// TIA Portal project "TestFineModuloPLC2SnideroEmanuele" (V19)

(* hardware
DEVICE "S7-1200 station_1"  S7-1200 Station
   slot 0: "Telaio di montaggio_0"  S7-1200 Rack  Rack  V1.0
   slot 1: "PLC_1"  CPU 1212C DC/DC/Rly  6ES7 212-1HE40-0XB0  V4.6
   slot 2: "DI 8/DQ 8x24VDC_1"  6ES7 223-1BH32-0XB0  V2.0
DEVICE "HMI_1"  KTP900 Basic PN
   slot 0: "HMI_1"  KTP900 Basic PN  6AV2 123-2JB03-0AX0  17.0.0.0
   slot 1: "HMI_RT_1"  KTP900 Basic PN  6AV2 123-2JB03-0AX0  17.0.0.0
   slot 5: "HMI_1.IE_CP_1"  PROFINET Interface  17.0.0.0
      slot 1: "Interfaccia_1 PROFINET"  PROFINET Interface
         slot 1: "Porta_1"  Port
DEVICE "SINAMICS G_1"  Sinamics.Device
   slot 0: "	_0"  Rail  SinamicsG120CRackP
   slot 0: "Drive_1"  G120C PN  6SL3210-1KE11-8AF2  4.7.14
      slot 1: "PROFINET interface"  MDD-SinamicsG120-P
      slot 3: "PM G120C"  PM G120C  6SL3210-1KE11-8AF2  -
*)

// ===== PLC "PLC_1"  CPU 1212C DC/DC/Rly =====

VAR_GLOBAL   // PLC tag table "Tabella delle variabili standard"
   "AbilitazioneAvvioNastro1" AT %I0.0 : Bool;
   "AbilitazioneAvvioNastro2" AT %I0.1 : Bool;
   "AbilitazioneAvvioNastro3" AT %I0.2 : Bool;
   "ArrestoNastro1" AT %I0.3 : Bool;
   "ArrestoNastro2" AT %I0.4 : Bool;
   "ArrestoNastro3" AT %I0.5 : Bool;
   "Emergenza" AT %I0.6 : Bool;
   "P01" AT %I0.7 : Bool;
   "P02" AT %I1.0 : Bool;
   "P1" AT %I1.1 : Bool;
   "P2" AT %I1.2 : Bool;
   "MotoreRobot" AT %Q0.0 : Bool;
   "MotoreAperturaPinza" AT %Q0.4 : Bool;
   "LEDLavorazione" AT %Q0.1 : Bool;
   "LEDRiposo" AT %Q0.2 : Bool;
   "LEDErrorePrelievoNastro1" AT %Q0.3 : Bool;
   "P03" AT %I1.4 : Bool;
   "P3" AT %I1.5 : Bool;
   "MotoreNastro1" AT %Q0.5 : Bool;
   "MotoreNastro2" AT %Q0.6 : Bool;
   "MotoreNastro3" AT %Q0.7 : Bool;
   "MotoreChiusuraPinza" AT %Q1.0 : Bool;
   "LEDErrorePrelievoNastro2" AT %Q1.1 : Bool;
   "Axis_1_Drive_IN" AT %I256.0 : "PD_TEL1_IN";
   "Axis_1_Drive_OUT" AT %Q256.0 : "PD_TEL1_OUT";
END_VAR

VAR_GLOBAL   // PLC tag table "Segnalazioni"
   "IndiceSegnalazioni" AT %MW100 : Int;
   "ErrorePrelievoNastro1" AT %M101.0 : Bool;
   "ErrorePrelievoNastro2" AT %M101.1 : Bool;
END_VAR

DATA_BLOCK "Sistema"   // DB1
{ S7_Optimized_Access := 'TRUE' }
VERSION : 0.1
   VAR
      DurataTrasportoNastri : Time := T#2500ms;
      DurataSpostamentoRobot : Time := T#2000ms;
      DurataMovimentoPinza : Time := T#2000ms;
      DurataPrelievoScatola : Time := T#20000ms;
      VolumeScatola : SInt := 6;
   END_VAR
   VAR RETAIN
      RiempimentoScatola : SInt;
   END_VAR
   VAR
      PP01 : Bool;
      PP02 : Bool;
      PP03 : Bool;
      PP1 : Bool;
      PP2 : Bool;
      PP3 : Bool;
      NMotoreNastro1 : Bool;
      NMotoreNastro2 : Bool;
      NMotoreNastro3 : Bool;
      NQTPSostituzioneScatola : Bool;
   END_VAR
   VAR RETAIN
      P1 : Bool;
      P2 : Bool;
   END_VAR
   VAR
      P3 : Bool;
      P03 : Bool;
      PP03Sistema : Bool;
      SetpointVelocitàNormato : Real;
   END_VAR
   VAR RETAIN
      SetpointVelocitàScalato : Real;
   END_VAR
BEGIN
END_DATA_BLOCK

DATA_BLOCK "HMI"   // DB4
{ S7_Optimized_Access := 'TRUE' }
VERSION : 0.1
   VAR
      StartNastro1 : Bool;
      StartNastro2 : Bool;
      StartNastro3 : Bool;
   END_VAR
   VAR RETAIN
      StopNastro1 : Bool := true;
      StopNastro2 : Bool := true;
      StopNastro3 : Bool := true;
      Emergenza : Bool;
   END_VAR
   VAR
      DitoFotocellulaNastro1 : Bool;
      DitoFotocellulaNastro2 : Bool;
      CaricamentoPezzoNastro1 : Bool;
      PCaricamentoPezzoNastro1 : Bool;
      CaricamentoPezzoNastro2 : Bool;
      PCaricamentoPezzoNastro2 : Bool;
   END_VAR
   VAR RETAIN
      Posizione1PinzaAperta : Bool;
      Posizione2PinzaAperta : Bool;
      Posizione3PinzaAperta : Bool;
      Posizione1PinzaChiusa : Bool;
      Posizione2PinzaChiusa : Bool;
      Posizione3PinzaChiusa : Bool;
      IndiceRicetta : Int := 1;
      NomeSetDati : String := 'Veloce';
   END_VAR
   VAR
      VisibilitàPezzoNastro1Veloce : Bool;
      VisibilitàPezzoNastro1Lento : Bool;
      VisibilitàPezzoNastro2Veloce : Bool;
      VisibilitàPezzoNastro2Lento : Bool;
      VisibilitàPezzoNastro3Veloce : Bool;
      VisibilitàPezzoNastro3Lento : Bool;
      SetpointVelocitàMotoreNastri : Real;
      VelocitàAttualeMotoreNastri : Real;
   END_VAR
BEGIN
END_DATA_BLOCK

DATA_BLOCK "Robot_DB"   // DB6
{ S7_Optimized_Access := 'TRUE' }
VERSION : 0.1
// stored: InstanceOfName Robot
"Robot"
BEGIN
END_DATA_BLOCK

DATA_BLOCK "SetDatiSistema"   // DB9
{ S7_Optimized_Access := 'TRUE' }
VERSION : 0.1
   VAR
      DurataTrasportoNastri : Time := T#5000ms;
      DurataSpostamentoRobot : Time := T#4000ms;
      VolumeScatola : SInt := 3;
   END_VAR
BEGIN
END_DATA_BLOCK

DATA_BLOCK "SetDatiSistemaVeloce"   // DB10
{ S7_Optimized_Access := 'TRUE' }
VERSION : 0.1
   VAR
      DurataTrasportoNastri : Time := T#5000ms;
      DurataSpostamentoRobot : Time := T#4000ms;
      VolumeScatola : SInt := 3;
   END_VAR
BEGIN
END_DATA_BLOCK

DATA_BLOCK "SetDatiSistemaLento"   // DB11
{ S7_Optimized_Access := 'TRUE' }
VERSION : 0.1
   VAR
      DurataTrasportoNastri : Time := T#5000ms;
      DurataSpostamentoRobot : Time := T#4000ms;
      VolumeScatola : SInt := 3;
   END_VAR
BEGIN
END_DATA_BLOCK

// folder: System blocks/Program resources

DATA_BLOCK "TPNastro1"   // DB2
{ S7_Optimized_Access := 'TRUE' }
AUTHOR : Simatic
FAMILY : IEC
NAME : IEC_TMR
VERSION : 1.0
// stored: InstanceOfName IEC_TIMER
"IEC_TIMER"
BEGIN
END_DATA_BLOCK

DATA_BLOCK "TPNastro2"   // DB3
{ S7_Optimized_Access := 'TRUE' }
AUTHOR : Simatic
FAMILY : IEC
NAME : IEC_TMR
VERSION : 1.0
// stored: InstanceOfName IEC_TIMER
"IEC_TIMER"
BEGIN
END_DATA_BLOCK

DATA_BLOCK "TPNastro3"   // DB5
{ S7_Optimized_Access := 'TRUE' }
AUTHOR : Simatic
FAMILY : IEC
NAME : IEC_TMR
VERSION : 1.0
// stored: InstanceOfName IEC_TIMER
"IEC_TIMER"
BEGIN
END_DATA_BLOCK

DATA_BLOCK "TPSostituzioneScatola"   // DB7
{ S7_Optimized_Access := 'TRUE' }
AUTHOR : Simatic
FAMILY : IEC
NAME : IEC_TMR
VERSION : 1.0
// stored: InstanceOfName IEC_TIMER
"IEC_TIMER"
BEGIN
END_DATA_BLOCK

// folder: (top level)

DATA_BLOCK "Axis_1"   // DB12, Motion_DB
{ S7_Optimized_Access := 'TRUE' }
AUTHOR : SIMATIC
FAMILY : BasicMC
NAME : TO_PosAx
VERSION : 8.0
// stored: InstanceOfName TO_PositioningAxis
"TO_PositioningAxis"
BEGIN
   // Axis.Drive.OfflineDataAdaption = TRUE
   // Axis.Drive.TelegramAddressOutCU = %Q256.0
   // Axis.Drive.TelegramAddressInCU = %I256.0
   // Axis.Drive.DoNameCU = Drive_1.Standard_telegram_1
   // Axis.Encoder.SelectedHscIndexCU = -1
   // Axis.LengthUnitNormalized.Time = 1
   // Axis.LengthUnitNormalized.Distance = -2
   // Axis.Encoder.DbTypeCU = Classic
   // Axis.Drive.DbTypeCU = Classic
END_DATA_BLOCK

FUNCTION_BLOCK "Robot"   // FB1, LAD
{ S7_Optimized_Access := 'TRUE' }
VERSION : 0.1
   VAR_INPUT
      Obiettivo : SInt;   // 0 = HOME, 1 = OK1, 2 = OK2, 3 = OK3
   END_VAR
   VAR RETAIN
      PosizioneAttuale : SInt;   // 0 = HOME, 1 = OK1, 2 = OK2, 3 = OK3
      PinzaAperta : Bool := true;
      PezzoPrelevatoDaNastro1 : Bool;
      PezzoPrelevatoDaNastro2 : Bool;
   END_VAR
   VAR
      TPRotazioneRobot : TP_TIME;
      NMotoreRobot : Bool;
      ObiettivoInRaggiungimento : SInt;
      PQTPRotazioneRobot : Bool;
      TPPinza : TP_TIME;
      NTPRotazioneRobot : Bool;
      NMotoreChiusuraPinza : Bool;
      NMotoreAperturaPinza : Bool;
      BloccoRotazione : Bool;
   END_VAR
   VAR_TEMP   // added for the SCL form of the ladder/FBD networks
      _w1 : Bool;
      _w2 : Bool;
      _w3 : Bool;
      _w4 : Bool;
      _w5 : Bool;
      _w6 : Bool;
      _w7 : Bool;
      _w8 : Bool;
   END_VAR
BEGIN

REGION Network 1
   // ROTAZIONE BRACCIO e APERTURA/CHIUSURA PINZA
   // 
   // L'input di posizione obiettivo può cambiare durante lo spostamento del robot, ma ciò non influisce sulla meta in raggiungimento.
   // Va però salvata la posizione in raggiugimento per la durata dello spostamento.
   // 
   // Prima di muovere verso la prossima posizione bisogna attendere eventuali manovre di pinza (a meno che non ci si trovi in HOME)
   // 
   // La pinza è inizialmente aperta e resta aperta dopo il deposito sul nastro 3
   // 
   // Le fotocellule di fine corsa dei nastri 1 e 2 vengono resettate automaticamente a fine operazione di prelievo. L'errore è simulabile tramite PLCSIM o apposito pulsante HMI.
   // 
   // Può accadere che venga premuto il pulsante di emergenza durante il movimento: in tal caso si arrestano i motori e, al termine dello scorrimento del tempo previsto per i loro azionamenti, si resetta il blocco rotativo
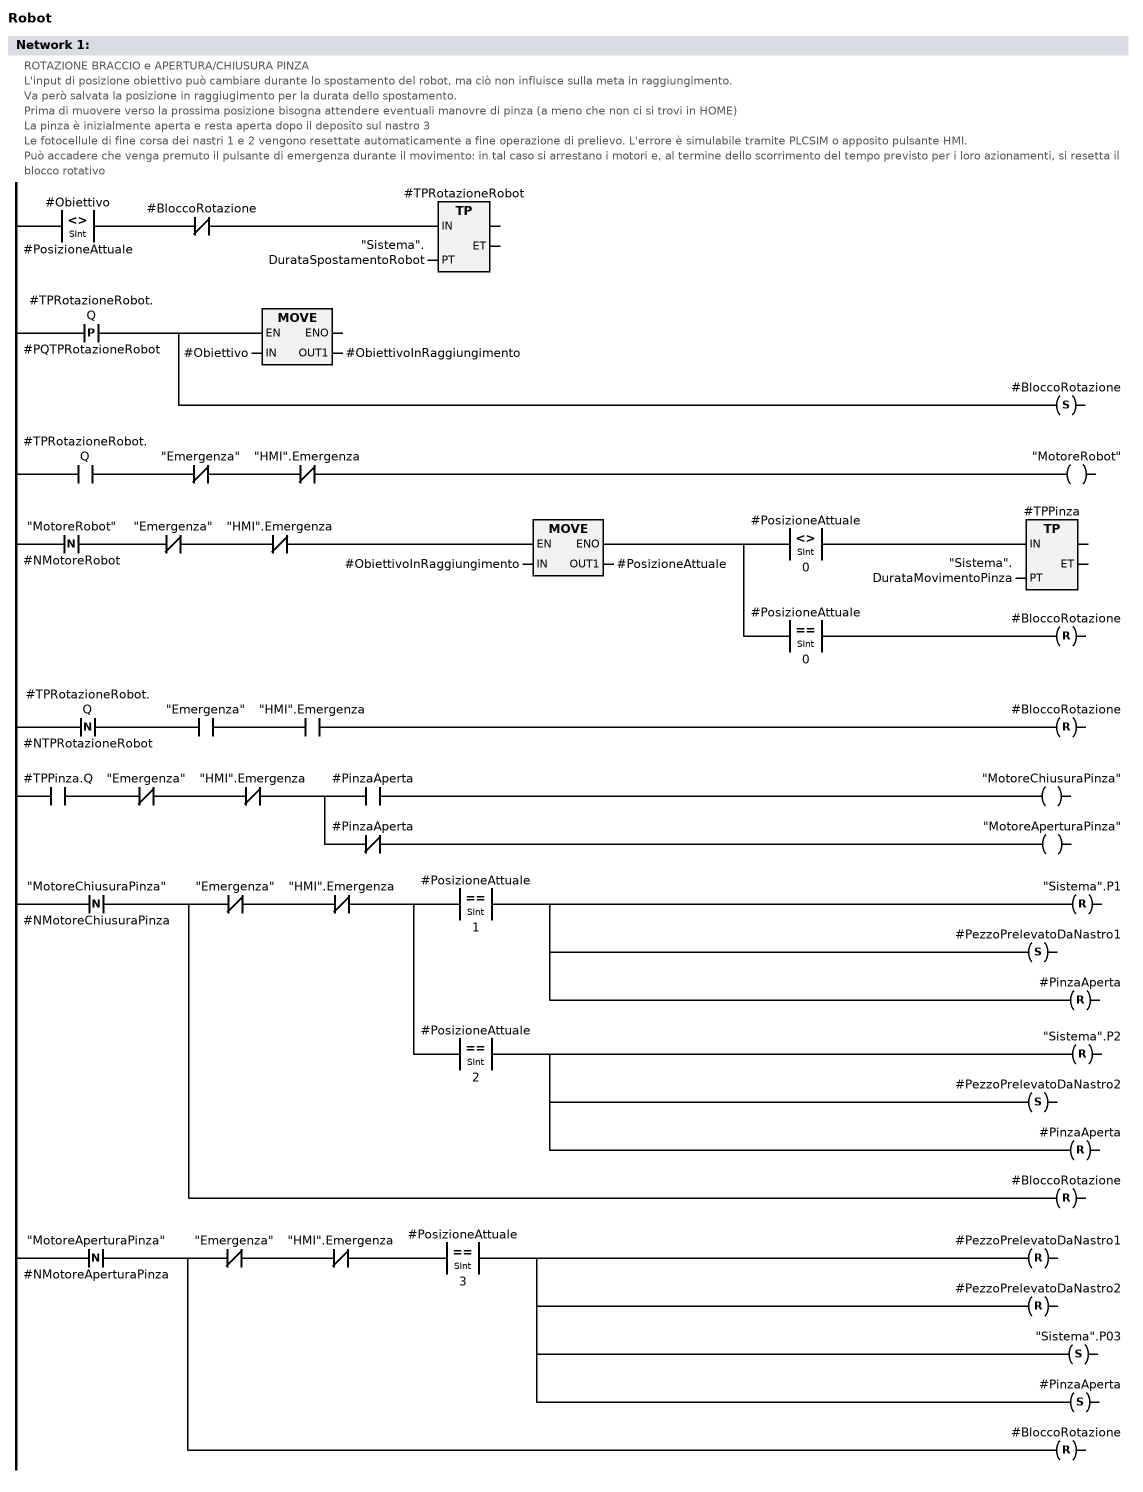
   #TPRotazioneRobot(IN := (#Obiettivo <> #PosizioneAttuale) AND NOT #BloccoRotazione,   // TP
                     PT := "Sistema".DurataSpostamentoRobot);
   #_w1 := #TPRotazioneRobot.Q AND NOT #PQTPRotazioneRobot;   // rising edge of #TPRotazioneRobot.Q
   #PQTPRotazioneRobot := #TPRotazioneRobot.Q;
   IF #_w1 THEN
       #ObiettivoInRaggiungimento := #Obiettivo;
       #BloccoRotazione := TRUE;
   END_IF;
   "MotoreRobot" := #TPRotazioneRobot.Q AND NOT "Emergenza" AND NOT "HMI".Emergenza;
   #_w2 := NOT "MotoreRobot" AND #NMotoreRobot;   // falling edge of "MotoreRobot"
   #NMotoreRobot := "MotoreRobot";
   #_w3 := #_w2 AND NOT "Emergenza" AND NOT "HMI".Emergenza;
   IF #_w3 THEN #PosizioneAttuale := #ObiettivoInRaggiungimento; END_IF;
   #TPPinza(IN := #_w3 AND (#PosizioneAttuale <> 0), PT := "Sistema".DurataMovimentoPinza);   // TP
   IF #_w3 AND (#PosizioneAttuale = 0) THEN #BloccoRotazione := FALSE; END_IF;
   #_w4 := NOT #TPRotazioneRobot.Q AND #NTPRotazioneRobot;   // falling edge of #TPRotazioneRobot.Q
   #NTPRotazioneRobot := #TPRotazioneRobot.Q;
   IF #_w4 AND "Emergenza" AND "HMI".Emergenza THEN #BloccoRotazione := FALSE; END_IF;
   #_w5 := #TPPinza.Q AND NOT "Emergenza" AND NOT "HMI".Emergenza;
   "MotoreChiusuraPinza" := #_w5 AND #PinzaAperta;
   "MotoreAperturaPinza" := #_w5 AND NOT #PinzaAperta;
   #_w6 := NOT "MotoreChiusuraPinza" AND #NMotoreChiusuraPinza;   // falling edge of "MotoreChiusuraPinza"
   #NMotoreChiusuraPinza := "MotoreChiusuraPinza";
   #_w7 := #_w6 AND NOT "Emergenza" AND NOT "HMI".Emergenza;
   IF #_w7 AND (#PosizioneAttuale = 1) THEN
       "Sistema".P1 := FALSE;
       #PezzoPrelevatoDaNastro1 := TRUE;
       #PinzaAperta := FALSE;
   END_IF;
   IF #_w7 AND (#PosizioneAttuale = 2) THEN
       "Sistema".P2 := FALSE;
       #PezzoPrelevatoDaNastro2 := TRUE;
       #PinzaAperta := FALSE;
   END_IF;
   IF #_w6 THEN #BloccoRotazione := FALSE; END_IF;
   #_w8 := NOT "MotoreAperturaPinza" AND #NMotoreAperturaPinza;   // falling edge of "MotoreAperturaPinza"
   #NMotoreAperturaPinza := "MotoreAperturaPinza";
   IF #_w8 AND NOT "Emergenza" AND NOT "HMI".Emergenza AND (#PosizioneAttuale = 3) THEN
       #PezzoPrelevatoDaNastro1 := FALSE;
       #PezzoPrelevatoDaNastro2 := FALSE;
       "Sistema".P03 := TRUE;
       #PinzaAperta := TRUE;
   END_IF;
   IF #_w8 THEN #BloccoRotazione := FALSE; END_IF;
END_REGION
END_FUNCTION_BLOCK

FUNCTION "AggiornamentoParametriRicetta" : Void   // FC2, LAD
{ S7_Optimized_Access := 'TRUE' }
VERSION : 0.1
   VAR_TEMP   // added for the SCL form of the ladder/FBD networks
      _w1 : Bool;
   END_VAR
BEGIN

REGION Network 1
   // Indice ricetta Sistema = 1
   // Indice salvato in Reciper Tag e in Data Record (HMI > Connections > Area Pointers)
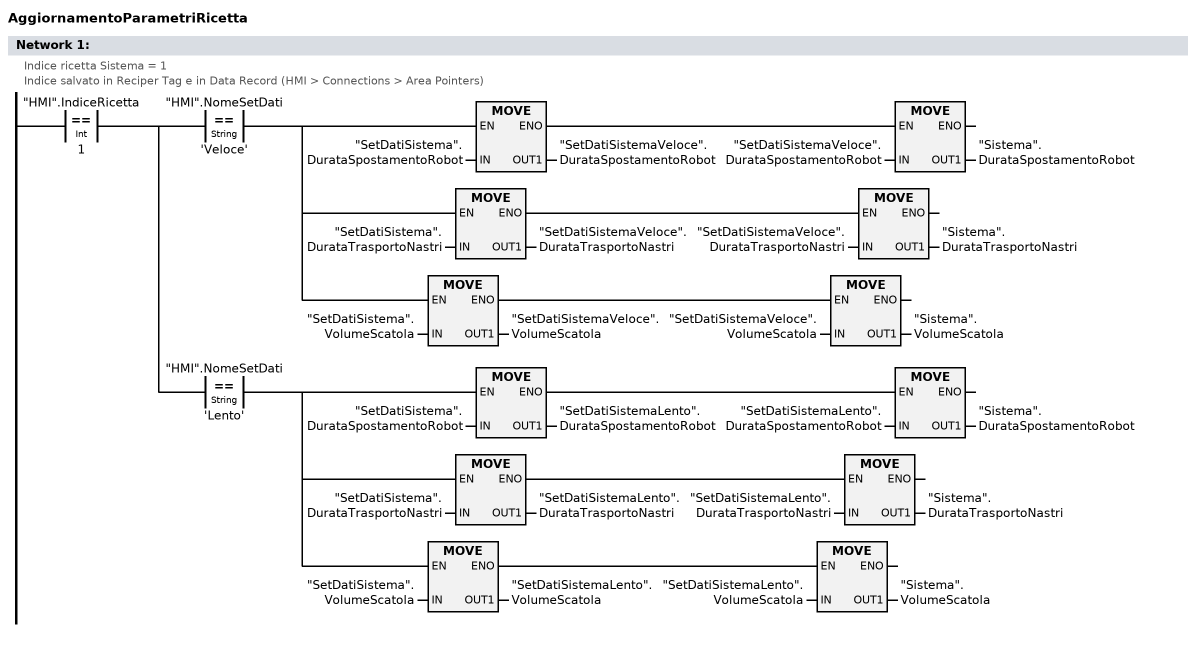
   RUNG wire#powerrail
      { S7_Templates := "SrcType := Int" } EQ_Contact(in1 := "HMI".IndiceRicetta, in2 := 1)
      wire#w1
      { S7_Templates := "SrcType := String" } EQ_Contact(in1 := "HMI".NomeSetDati, in2 := 'Veloce')
      wire#w2
      Move(in := "SetDatiSistema".DurataSpostamentoRobot, out1 => "SetDatiSistemaVeloce".DurataSpostamentoRobot)
      Move(in := "SetDatiSistemaVeloce".DurataSpostamentoRobot, out1 => "Sistema".DurataSpostamentoRobot)
   END_RUNG
   RUNG wire#w2
      Move(in := "SetDatiSistema".DurataTrasportoNastri, out1 => "SetDatiSistemaVeloce".DurataTrasportoNastri)
      Move(in := "SetDatiSistemaVeloce".DurataTrasportoNastri, out1 => "Sistema".DurataTrasportoNastri)
   END_RUNG
   RUNG wire#w2
      Move(in := "SetDatiSistema".VolumeScatola, out1 => "SetDatiSistemaVeloce".VolumeScatola)
      Move(in := "SetDatiSistemaVeloce".VolumeScatola, out1 => "Sistema".VolumeScatola)
   END_RUNG
   RUNG wire#w1
      { S7_Templates := "SrcType := String" } EQ_Contact(in1 := "HMI".NomeSetDati, in2 := 'Lento')
      wire#w3
      Move(in := "SetDatiSistema".DurataSpostamentoRobot, out1 => "SetDatiSistemaLento".DurataSpostamentoRobot)
      Move(in := "SetDatiSistemaLento".DurataSpostamentoRobot, out1 => "Sistema".DurataSpostamentoRobot)
   END_RUNG
   RUNG wire#w3
      Move(in := "SetDatiSistema".DurataTrasportoNastri, out1 => "SetDatiSistemaLento".DurataTrasportoNastri)
      Move(in := "SetDatiSistemaLento".DurataTrasportoNastri, out1 => "Sistema".DurataTrasportoNastri)
   END_RUNG
   RUNG wire#w3
      Move(in := "SetDatiSistema".VolumeScatola, out1 => "SetDatiSistemaLento".VolumeScatola)
      Move(in := "SetDatiSistemaLento".VolumeScatola, out1 => "Sistema".VolumeScatola)
   END_RUNG
   // the same network as SCL:
   #_w1 := "HMI".IndiceRicetta = 1;
   IF #_w1 AND ("HMI".NomeSetDati = 'Veloce') THEN
       "SetDatiSistemaVeloce".DurataSpostamentoRobot := "SetDatiSistema".DurataSpostamentoRobot;
       "Sistema".DurataSpostamentoRobot := "SetDatiSistemaVeloce".DurataSpostamentoRobot;
       "SetDatiSistemaVeloce".DurataTrasportoNastri := "SetDatiSistema".DurataTrasportoNastri;
       "Sistema".DurataTrasportoNastri := "SetDatiSistemaVeloce".DurataTrasportoNastri;
       "SetDatiSistemaVeloce".VolumeScatola := "SetDatiSistema".VolumeScatola;
       "Sistema".VolumeScatola := "SetDatiSistemaVeloce".VolumeScatola;
   END_IF;
   IF #_w1 AND ("HMI".NomeSetDati = 'Lento') THEN
       "SetDatiSistemaLento".DurataSpostamentoRobot := "SetDatiSistema".DurataSpostamentoRobot;
       "Sistema".DurataSpostamentoRobot := "SetDatiSistemaLento".DurataSpostamentoRobot;
       "SetDatiSistemaLento".DurataTrasportoNastri := "SetDatiSistema".DurataTrasportoNastri;
       "Sistema".DurataTrasportoNastri := "SetDatiSistemaLento".DurataTrasportoNastri;
       "SetDatiSistemaLento".VolumeScatola := "SetDatiSistema".VolumeScatola;
       "Sistema".VolumeScatola := "SetDatiSistemaLento".VolumeScatola;
   END_IF;
END_REGION
END_FUNCTION

ORGANIZATION_BLOCK "Main"   // OB1, LAD, ProgramCycle
TITLE = "Main Program Sweep (Cycle)"
{ S7_Optimized_Access := 'TRUE' }
VERSION : 0.1
   VAR_INPUT
      Initial_Call : Bool;   // Initial call of this OB
      Remanence : Bool;   // =True, if remanent data are available
   END_VAR
   VAR_TEMP   // added for the SCL form of the ladder/FBD networks
      _w1 : Bool;
      _w2 : Bool;
      _w3 : Bool;
      _w4 : Bool;
   END_VAR
BEGIN

REGION Network 1
   // Trasporto pezzi nastro 1
   // 
   // Non è possibile posizionare pezzi sui nastri finché ne sono in trasporto altri (o, meglio, è possibile ma il motore si fermerà si muoverà solamente per permettere) o la fotocellula di fine corsa non viene liberata (il motore non si aziona)
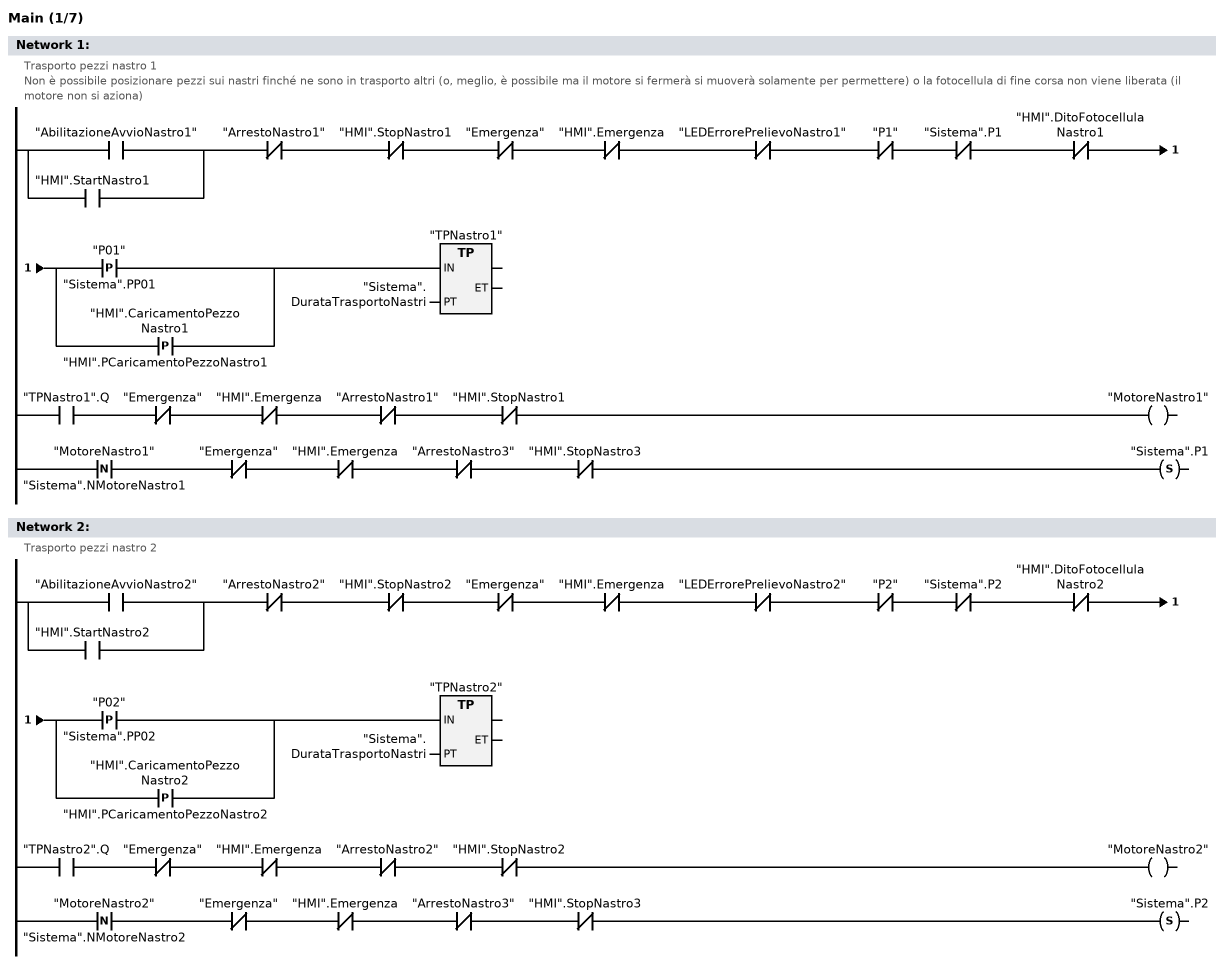
   #_w1 := ("AbilitazioneAvvioNastro1" OR "HMI".StartNastro1) AND NOT "ArrestoNastro1" AND NOT "HMI".StopNastro1 AND NOT "Emergenza" AND NOT "HMI".Emergenza AND NOT "LEDErrorePrelievoNastro1" AND NOT "P1" AND NOT "Sistema".P1 AND NOT "HMI".DitoFotocellulaNastro1 AND "P01" AND NOT "Sistema".PP01;   // rising edge of "P01"
   "Sistema".PP01 := "P01";
   #_w2 := ("AbilitazioneAvvioNastro1" OR "HMI".StartNastro1) AND NOT "ArrestoNastro1" AND NOT "HMI".StopNastro1 AND NOT "Emergenza" AND NOT "HMI".Emergenza AND NOT "LEDErrorePrelievoNastro1" AND NOT "P1" AND NOT "Sistema".P1 AND NOT "HMI".DitoFotocellulaNastro1 AND "HMI".CaricamentoPezzoNastro1 AND NOT "HMI".PCaricamentoPezzoNastro1;   // rising edge of "HMI".CaricamentoPezzoNastro1
   "HMI".PCaricamentoPezzoNastro1 := "HMI".CaricamentoPezzoNastro1;
   "TPNastro1".TP(IN := #_w1 OR #_w2, PT := "Sistema".DurataTrasportoNastri);
   "MotoreNastro1" := "TPNastro1".Q AND NOT "Emergenza" AND NOT "HMI".Emergenza AND NOT "ArrestoNastro1" AND NOT "HMI".StopNastro1;
   #_w3 := NOT "MotoreNastro1" AND "Sistema".NMotoreNastro1;   // falling edge of "MotoreNastro1"
   "Sistema".NMotoreNastro1 := "MotoreNastro1";
   IF #_w3 AND NOT "Emergenza" AND NOT "HMI".Emergenza AND NOT "ArrestoNastro3" AND NOT "HMI".StopNastro3 THEN
       "Sistema".P1 := TRUE;
   END_IF;
END_REGION

REGION Network 2
   // Trasporto pezzi nastro 2
   #_w1 := ("AbilitazioneAvvioNastro2" OR "HMI".StartNastro2) AND NOT "ArrestoNastro2" AND NOT "HMI".StopNastro2 AND NOT "Emergenza" AND NOT "HMI".Emergenza AND NOT "LEDErrorePrelievoNastro2" AND NOT "P2" AND NOT "Sistema".P2 AND NOT "HMI".DitoFotocellulaNastro2 AND "P02" AND NOT "Sistema".PP02;   // rising edge of "P02"
   "Sistema".PP02 := "P02";
   #_w2 := ("AbilitazioneAvvioNastro2" OR "HMI".StartNastro2) AND NOT "ArrestoNastro2" AND NOT "HMI".StopNastro2 AND NOT "Emergenza" AND NOT "HMI".Emergenza AND NOT "LEDErrorePrelievoNastro2" AND NOT "P2" AND NOT "Sistema".P2 AND NOT "HMI".DitoFotocellulaNastro2 AND "HMI".CaricamentoPezzoNastro2 AND NOT "HMI".PCaricamentoPezzoNastro2;   // rising edge of "HMI".CaricamentoPezzoNastro2
   "HMI".PCaricamentoPezzoNastro2 := "HMI".CaricamentoPezzoNastro2;
   "TPNastro2".TP(IN := #_w1 OR #_w2, PT := "Sistema".DurataTrasportoNastri);
   "MotoreNastro2" := "TPNastro2".Q AND NOT "Emergenza" AND NOT "HMI".Emergenza AND NOT "ArrestoNastro2" AND NOT "HMI".StopNastro2;
   #_w3 := NOT "MotoreNastro2" AND "Sistema".NMotoreNastro2;   // falling edge of "MotoreNastro2"
   "Sistema".NMotoreNastro2 := "MotoreNastro2";
   IF #_w3 AND NOT "Emergenza" AND NOT "HMI".Emergenza AND NOT "ArrestoNastro3" AND NOT "HMI".StopNastro3 THEN
       "Sistema".P2 := TRUE;
   END_IF;
END_REGION

REGION Network 3
   // Trasporto pezzi nastro 3 e riempimento scatola
   // 
   // Il nastro 3 non si muove se la scatola piena non è stata rimpiazzata
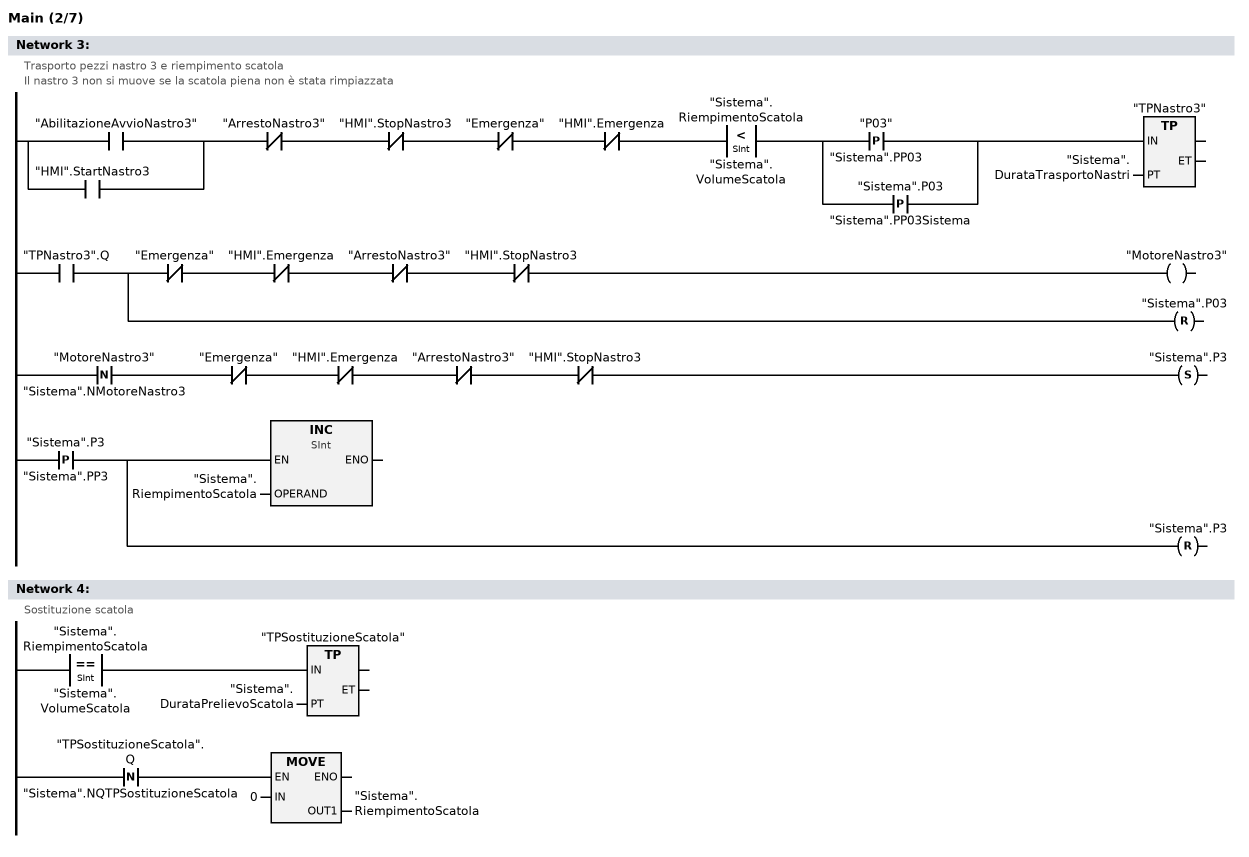
   #_w1 := ("AbilitazioneAvvioNastro3" OR "HMI".StartNastro3) AND NOT "ArrestoNastro3" AND NOT "HMI".StopNastro3 AND NOT "Emergenza" AND NOT "HMI".Emergenza AND ("Sistema".RiempimentoScatola < "Sistema".VolumeScatola) AND "P03" AND NOT "Sistema".PP03;   // rising edge of "P03"
   "Sistema".PP03 := "P03";
   #_w2 := ("AbilitazioneAvvioNastro3" OR "HMI".StartNastro3) AND NOT "ArrestoNastro3" AND NOT "HMI".StopNastro3 AND NOT "Emergenza" AND NOT "HMI".Emergenza AND ("Sistema".RiempimentoScatola < "Sistema".VolumeScatola) AND "Sistema".P03 AND NOT "Sistema".PP03Sistema;   // rising edge of "Sistema".P03
   "Sistema".PP03Sistema := "Sistema".P03;
   "TPNastro3".TP(IN := #_w1 OR #_w2, PT := "Sistema".DurataTrasportoNastri);
   "MotoreNastro3" := "TPNastro3".Q AND NOT "Emergenza" AND NOT "HMI".Emergenza AND NOT "ArrestoNastro3" AND NOT "HMI".StopNastro3;
   IF "TPNastro3".Q THEN "Sistema".P03 := FALSE; END_IF;
   #_w3 := NOT "MotoreNastro3" AND "Sistema".NMotoreNastro3;   // falling edge of "MotoreNastro3"
   "Sistema".NMotoreNastro3 := "MotoreNastro3";
   IF #_w3 AND NOT "Emergenza" AND NOT "HMI".Emergenza AND NOT "ArrestoNastro3" AND NOT "HMI".StopNastro3 THEN
       "Sistema".P3 := TRUE;
   END_IF;
   #_w4 := "Sistema".P3 AND NOT "Sistema".PP3;   // rising edge of "Sistema".P3
   "Sistema".PP3 := "Sistema".P3;
   IF #_w4 THEN
       "Sistema".RiempimentoScatola := "Sistema".RiempimentoScatola + 1;
       "Sistema".P3 := FALSE;
   END_IF;
END_REGION

REGION Network 4
   // Sostituzione scatola
   "TPSostituzioneScatola".TP(IN := "Sistema".RiempimentoScatola = "Sistema".VolumeScatola,
                           PT := "Sistema".DurataPrelievoScatola);
   #_w1 := NOT "TPSostituzioneScatola".Q AND "Sistema".NQTPSostituzioneScatola;   // falling edge of "TPSostituzioneScatola".Q
   "Sistema".NQTPSostituzioneScatola := "TPSostituzioneScatola".Q;
   IF #_w1 THEN "Sistema".RiempimentoScatola := 0; END_IF;
END_REGION

REGION Network 5
   // MOVIMENTAZIONE ROBOT
   // 
   // Spostamenti
   // - home => nastro 1/2
   // - nastro 1/2 => nastro 3
   // - nastro 3 => nastro1/2/home (se assenti pezzi da prelevare)
   // 
   // L'oggetto non viene prelevato per essere rilasciato sul nastro 3 finché il motore del nastro è in stato di arresto o la scatola è piena
   // Può però essere prelevato se il nastro 3 è in movimento perché vi è tempo sufficiente a completare l'inscatolamento del precedente prima che venga rilasciato.
   // 
   // Il nastro 1 ha precedenza sul 2
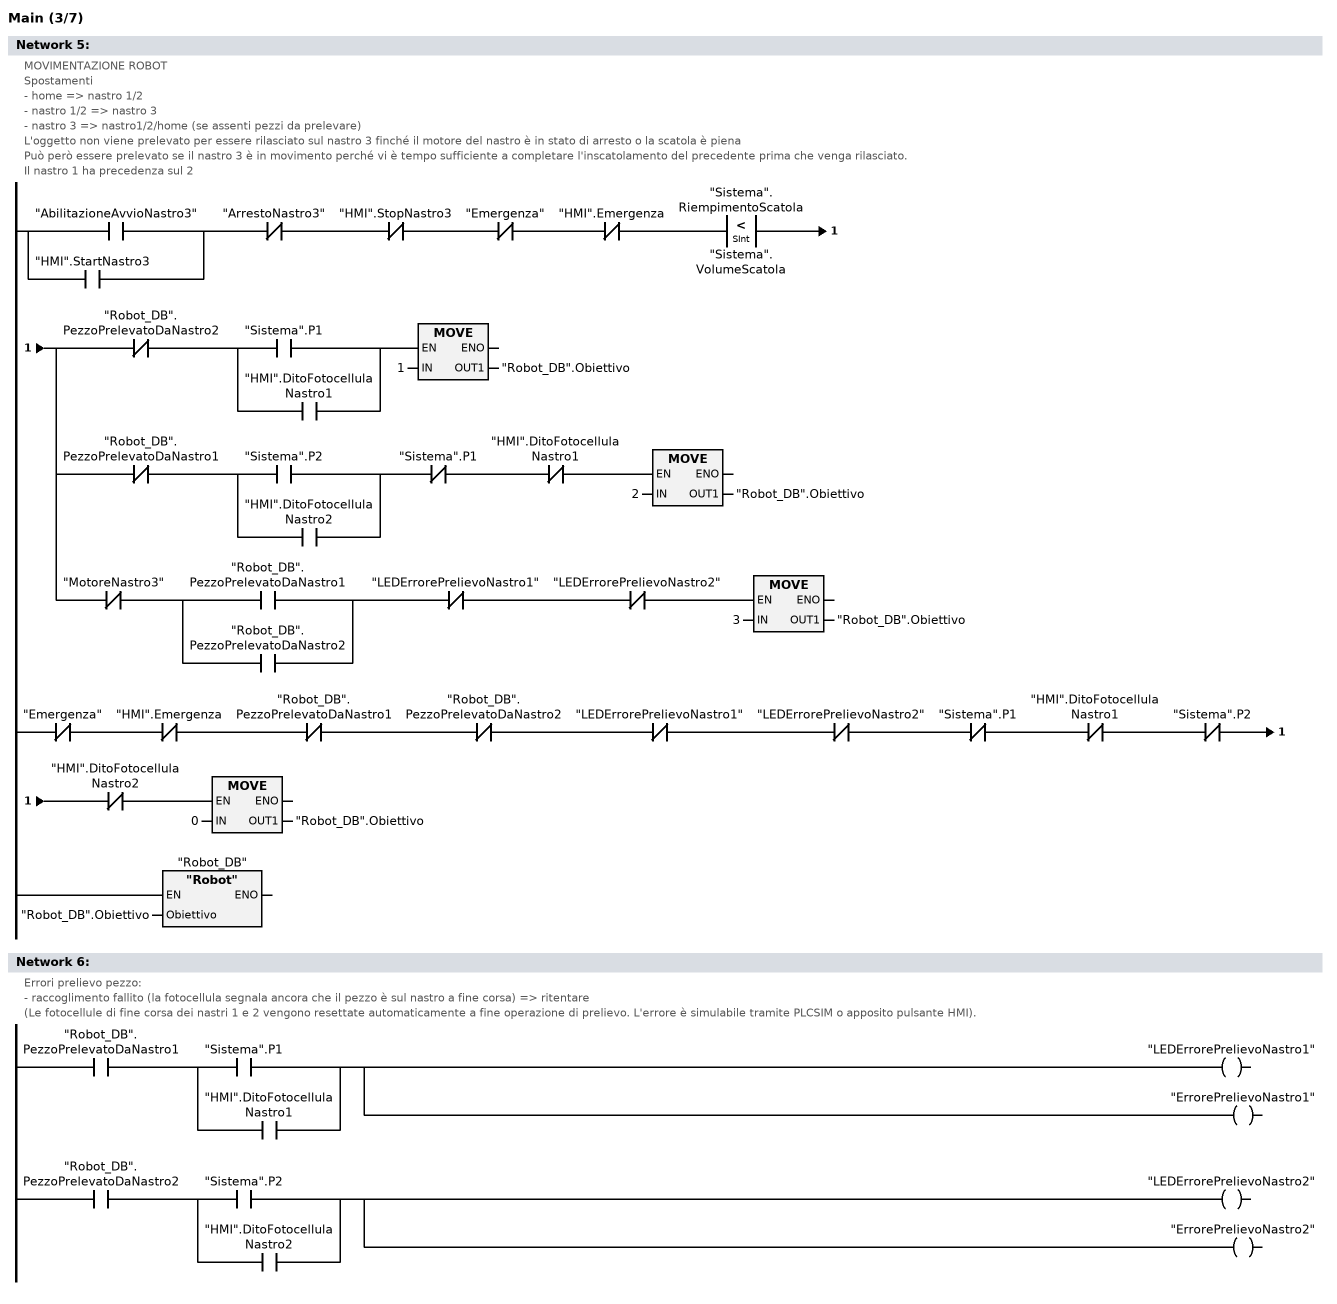
   RUNG wire#powerrail
      Contact( "AbilitazioneAvvioNastro3" )
      wire#w1
      I_Contact( "ArrestoNastro3" )
      I_Contact( "HMI".StopNastro3 )
      I_Contact( "Emergenza" )
      I_Contact( "HMI".Emergenza )
      { S7_Templates := "SrcType := SInt" } LT_Contact(in1 := "Sistema".RiempimentoScatola, in2 := "Sistema".VolumeScatola)
      wire#w2
      I_Contact( "Robot_DB".PezzoPrelevatoDaNastro2 )
      wire#w3
      Contact( "Sistema".P1 )
      wire#w4
      Move(in := 1, out1 => "Robot_DB".Obiettivo)
   END_RUNG
   RUNG wire#powerrail
      Contact( "HMI".StartNastro3 )
   END_RUNG wire#w1
   RUNG wire#w3
      Contact( "HMI".DitoFotocellulaNastro1 )
   END_RUNG wire#w4
   RUNG wire#w2
      I_Contact( "Robot_DB".PezzoPrelevatoDaNastro1 )
      wire#w5
      Contact( "Sistema".P2 )
      wire#w6
      I_Contact( "Sistema".P1 )
      I_Contact( "HMI".DitoFotocellulaNastro1 )
      Move(in := 2, out1 => "Robot_DB".Obiettivo)
   END_RUNG
   RUNG wire#w5
      Contact( "HMI".DitoFotocellulaNastro2 )
   END_RUNG wire#w6
   RUNG wire#w2
      I_Contact( "MotoreNastro3" )
      wire#w7
      Contact( "Robot_DB".PezzoPrelevatoDaNastro1 )
      wire#w8
      I_Contact( "LEDErrorePrelievoNastro1" )
      I_Contact( "LEDErrorePrelievoNastro2" )
      Move(in := 3, out1 => "Robot_DB".Obiettivo)
   END_RUNG
   RUNG wire#w7
      Contact( "Robot_DB".PezzoPrelevatoDaNastro2 )
   END_RUNG wire#w8
   RUNG wire#powerrail
      I_Contact( "Emergenza" )
      I_Contact( "HMI".Emergenza )
      I_Contact( "Robot_DB".PezzoPrelevatoDaNastro1 )
      I_Contact( "Robot_DB".PezzoPrelevatoDaNastro2 )
      I_Contact( "LEDErrorePrelievoNastro1" )
      I_Contact( "LEDErrorePrelievoNastro2" )
      I_Contact( "Sistema".P1 )
      I_Contact( "HMI".DitoFotocellulaNastro1 )
      I_Contact( "Sistema".P2 )
      I_Contact( "HMI".DitoFotocellulaNastro2 )
      Move(in := 0, out1 => "Robot_DB".Obiettivo)
   END_RUNG
   RUNG wire#powerrail
      "Robot_DB"(Obiettivo := "Robot_DB".Obiettivo)
   END_RUNG
   // the same network as SCL:
   #_w1 := ("AbilitazioneAvvioNastro3" OR "HMI".StartNastro3) AND NOT "ArrestoNastro3" AND NOT "HMI".StopNastro3 AND NOT "Emergenza" AND NOT "HMI".Emergenza AND ("Sistema".RiempimentoScatola < "Sistema".VolumeScatola);
   IF #_w1 AND NOT "Robot_DB".PezzoPrelevatoDaNastro2 AND ("Sistema".P1 OR "HMI".DitoFotocellulaNastro1) THEN
       "Robot_DB".Obiettivo := 1;
   END_IF;
   IF #_w1 AND NOT "Robot_DB".PezzoPrelevatoDaNastro1 AND ("Sistema".P2 OR "HMI".DitoFotocellulaNastro2) AND NOT "Sistema".P1 AND NOT "HMI".DitoFotocellulaNastro1 THEN
       "Robot_DB".Obiettivo := 2;
   END_IF;
   IF #_w1 AND NOT "MotoreNastro3" AND ("Robot_DB".PezzoPrelevatoDaNastro1 OR "Robot_DB".PezzoPrelevatoDaNastro2) AND NOT "LEDErrorePrelievoNastro1" AND NOT "LEDErrorePrelievoNastro2" THEN
       "Robot_DB".Obiettivo := 3;
   END_IF;
   IF NOT "Emergenza" AND NOT "HMI".Emergenza AND NOT "Robot_DB".PezzoPrelevatoDaNastro1 AND NOT "Robot_DB".PezzoPrelevatoDaNastro2 AND NOT "LEDErrorePrelievoNastro1" AND NOT "LEDErrorePrelievoNastro2" AND NOT "Sistema".P1 AND NOT "HMI".DitoFotocellulaNastro1 AND NOT "Sistema".P2 AND NOT "HMI".DitoFotocellulaNastro2 THEN
       "Robot_DB".Obiettivo := 0;
   END_IF;
   "Robot_DB"(Obiettivo := "Robot_DB".Obiettivo);   // "Robot"
END_REGION

REGION Network 6
   // Errori prelievo pezzo: 
   // - raccoglimento fallito (la fotocellula segnala ancora che il pezzo è sul nastro a fine corsa) => ritentare
   // 
   // (Le fotocellule di fine corsa dei nastri 1 e 2 vengono resettate automaticamente a fine operazione di prelievo. L'errore è simulabile tramite PLCSIM o apposito pulsante HMI).
   RUNG wire#powerrail
      Contact( "Robot_DB".PezzoPrelevatoDaNastro1 )
      wire#w1
      Contact( "Sistema".P1 )
      wire#w2
      Coil( "LEDErrorePrelievoNastro1" )
   END_RUNG
   RUNG wire#w1
      Contact( "HMI".DitoFotocellulaNastro1 )
   END_RUNG wire#w2
   RUNG wire#w2
      Coil( "ErrorePrelievoNastro1" )
   END_RUNG
   RUNG wire#powerrail
      Contact( "Robot_DB".PezzoPrelevatoDaNastro2 )
      wire#w3
      Contact( "Sistema".P2 )
      wire#w4
      Coil( "LEDErrorePrelievoNastro2" )
   END_RUNG
   RUNG wire#w3
      Contact( "HMI".DitoFotocellulaNastro2 )
   END_RUNG wire#w4
   RUNG wire#w4
      Coil( "ErrorePrelievoNastro2" )
   END_RUNG
   // the same network as SCL:
   "LEDErrorePrelievoNastro1" := "Robot_DB".PezzoPrelevatoDaNastro1 AND ("Sistema".P1 OR "HMI".DitoFotocellulaNastro1);
   "ErrorePrelievoNastro1" := "LEDErrorePrelievoNastro1";
   "LEDErrorePrelievoNastro2" := "Robot_DB".PezzoPrelevatoDaNastro2 AND ("Sistema".P2 OR "HMI".DitoFotocellulaNastro2);
   "ErrorePrelievoNastro2" := "LEDErrorePrelievoNastro2";
END_REGION

REGION Network 7
   // Alimentazione LED marcia sistema quando:
   // - il robot è in rotazione o in azionamento pinza
   // - un nastro è in scorrimento
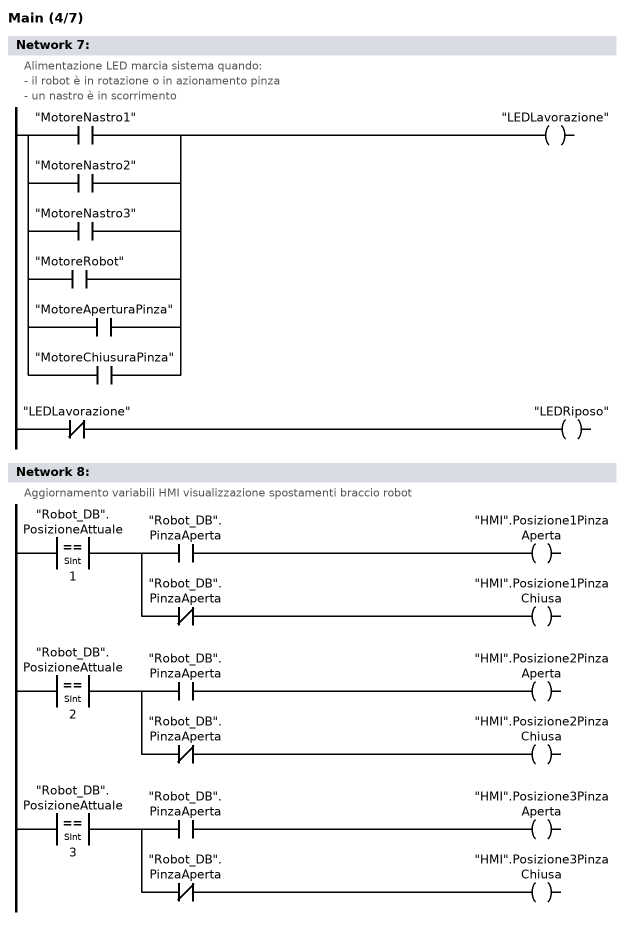
   RUNG wire#powerrail
      Contact( "MotoreNastro1" )
      wire#w1
      Coil( "LEDLavorazione" )
   END_RUNG
   RUNG wire#powerrail
      Contact( "MotoreNastro2" )
   END_RUNG wire#w1
   RUNG wire#powerrail
      Contact( "MotoreNastro3" )
   END_RUNG wire#w1
   RUNG wire#powerrail
      Contact( "MotoreRobot" )
   END_RUNG wire#w1
   RUNG wire#powerrail
      Contact( "MotoreAperturaPinza" )
   END_RUNG wire#w1
   RUNG wire#powerrail
      Contact( "MotoreChiusuraPinza" )
   END_RUNG wire#w1
   RUNG wire#powerrail
      I_Contact( "LEDLavorazione" )
      Coil( "LEDRiposo" )
   END_RUNG
   // the same network as SCL:
   "LEDLavorazione" := "MotoreNastro1" OR "MotoreNastro2" OR "MotoreNastro3" OR "MotoreRobot" OR "MotoreAperturaPinza" OR "MotoreChiusuraPinza";
   "LEDRiposo" := NOT "LEDLavorazione";
END_REGION

REGION Network 8
   // Aggiornamento variabili HMI visualizzazione spostamenti braccio robot
   RUNG wire#powerrail
      { S7_Templates := "SrcType := SInt" } EQ_Contact(in1 := "Robot_DB".PosizioneAttuale, in2 := 1)
      wire#w1
      Contact( "Robot_DB".PinzaAperta )
      Coil( "HMI".Posizione1PinzaAperta )
   END_RUNG
   RUNG wire#w1
      I_Contact( "Robot_DB".PinzaAperta )
      Coil( "HMI".Posizione1PinzaChiusa )
   END_RUNG
   RUNG wire#powerrail
      { S7_Templates := "SrcType := SInt" } EQ_Contact(in1 := "Robot_DB".PosizioneAttuale, in2 := 2)
      wire#w2
      Contact( "Robot_DB".PinzaAperta )
      Coil( "HMI".Posizione2PinzaAperta )
   END_RUNG
   RUNG wire#w2
      I_Contact( "Robot_DB".PinzaAperta )
      Coil( "HMI".Posizione2PinzaChiusa )
   END_RUNG
   RUNG wire#powerrail
      { S7_Templates := "SrcType := SInt" } EQ_Contact(in1 := "Robot_DB".PosizioneAttuale, in2 := 3)
      wire#w3
      Contact( "Robot_DB".PinzaAperta )
      Coil( "HMI".Posizione3PinzaAperta )
   END_RUNG
   RUNG wire#w3
      I_Contact( "Robot_DB".PinzaAperta )
      Coil( "HMI".Posizione3PinzaChiusa )
   END_RUNG
   // the same network as SCL:
   #_w1 := "Robot_DB".PosizioneAttuale = 1;
   "HMI".Posizione1PinzaAperta := #_w1 AND "Robot_DB".PinzaAperta;
   "HMI".Posizione1PinzaChiusa := #_w1 AND NOT "Robot_DB".PinzaAperta;
   #_w2 := "Robot_DB".PosizioneAttuale = 2;
   "HMI".Posizione2PinzaAperta := #_w2 AND "Robot_DB".PinzaAperta;
   "HMI".Posizione2PinzaChiusa := #_w2 AND NOT "Robot_DB".PinzaAperta;
   #_w3 := "Robot_DB".PosizioneAttuale = 3;
   "HMI".Posizione3PinzaAperta := #_w3 AND "Robot_DB".PinzaAperta;
   "HMI".Posizione3PinzaChiusa := #_w3 AND NOT "Robot_DB".PinzaAperta;
END_REGION

REGION Network 9
   // Aggiornamento variabili HMI visualizzazione pezzi in movimento sui nastri
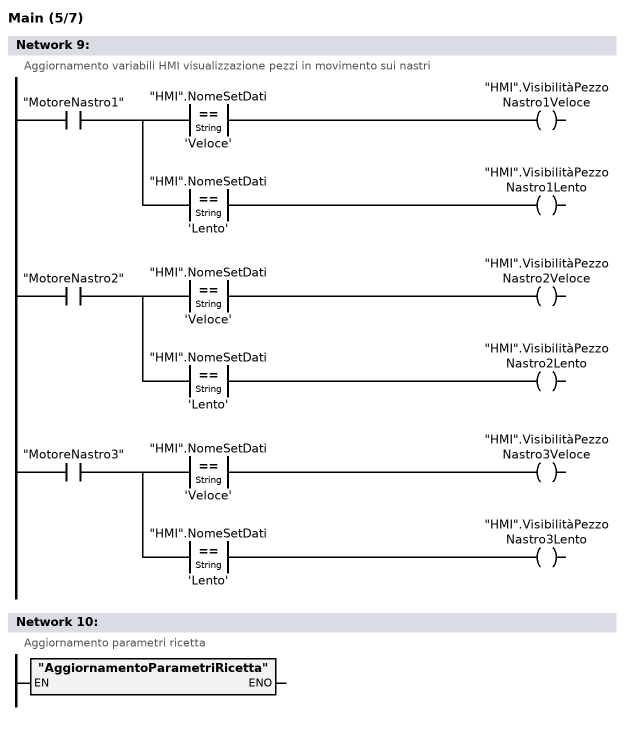
   RUNG wire#powerrail
      Contact( "MotoreNastro1" )
      wire#w1
      { S7_Templates := "SrcType := String" } EQ_Contact(in1 := "HMI".NomeSetDati, in2 := 'Veloce')
      Coil( "HMI".VisibilitàPezzoNastro1Veloce )
   END_RUNG
   RUNG wire#w1
      { S7_Templates := "SrcType := String" } EQ_Contact(in1 := "HMI".NomeSetDati, in2 := 'Lento')
      Coil( "HMI".VisibilitàPezzoNastro1Lento )
   END_RUNG
   RUNG wire#powerrail
      Contact( "MotoreNastro2" )
      wire#w2
      { S7_Templates := "SrcType := String" } EQ_Contact(in1 := "HMI".NomeSetDati, in2 := 'Veloce')
      Coil( "HMI".VisibilitàPezzoNastro2Veloce )
   END_RUNG
   RUNG wire#w2
      { S7_Templates := "SrcType := String" } EQ_Contact(in1 := "HMI".NomeSetDati, in2 := 'Lento')
      Coil( "HMI".VisibilitàPezzoNastro2Lento )
   END_RUNG
   RUNG wire#powerrail
      Contact( "MotoreNastro3" )
      wire#w3
      { S7_Templates := "SrcType := String" } EQ_Contact(in1 := "HMI".NomeSetDati, in2 := 'Veloce')
      Coil( "HMI".VisibilitàPezzoNastro3Veloce )
   END_RUNG
   RUNG wire#w3
      { S7_Templates := "SrcType := String" } EQ_Contact(in1 := "HMI".NomeSetDati, in2 := 'Lento')
      Coil( "HMI".VisibilitàPezzoNastro3Lento )
   END_RUNG
   // the same network as SCL:
   "HMI".VisibilitàPezzoNastro1Veloce := "MotoreNastro1" AND ("HMI".NomeSetDati = 'Veloce');
   "HMI".VisibilitàPezzoNastro1Lento := "MotoreNastro1" AND ("HMI".NomeSetDati = 'Lento');
   "HMI".VisibilitàPezzoNastro2Veloce := "MotoreNastro2" AND ("HMI".NomeSetDati = 'Veloce');
   "HMI".VisibilitàPezzoNastro2Lento := "MotoreNastro2" AND ("HMI".NomeSetDati = 'Lento');
   "HMI".VisibilitàPezzoNastro3Veloce := "MotoreNastro3" AND ("HMI".NomeSetDati = 'Veloce');
   "HMI".VisibilitàPezzoNastro3Lento := "MotoreNastro3" AND ("HMI".NomeSetDati = 'Lento');
END_REGION

REGION Network 10
   // Aggiornamento parametri ricetta
   RUNG wire#powerrail
      "AggiornamentoParametriRicetta"()
   END_RUNG
   // the same network as SCL:
   "AggiornamentoParametriRicetta"();
END_REGION

REGION Network 11: 0-->1; 1 = Enable the drive (OFF2 / OFF 3 are 1 in default status) (OFF1 = 0-->1)
   // Regolazione (su base ricetta) velocità motore nastri con FB SINAMICS (calcolo lato drive)
   // 
   // Parametri driver
   // - Rated speed (parametro p(0)311) = Velocità nominale motore (velocità di coppia nominale) = velocità di sincronismo x (1 - scorrimento a pieno carico)
   // - Reference speed (p2000) = massima velocità di riferimento scalare telegramma (consigliato eguagliare a Maximum speed: se le eccede il driver non supera comunque MaximumSpeed)
   // - Maximum speed (p1082) = velocità (sicura) massima motore
   // 
   // Nel progetto il movimento "veloce" del motore è a velocità nominale (come settato nel driver)
   // 
   // Parametri SinaSpeed lavorando con telegramma tipo 1 (SinaPos lavora invece con 111, supportato solo dai driver con interfacciamento encoder integrato)
   // - Refspeed = riferimento scalatura velocità telegramma (parametro p2000 del driver)
   // - ConfigAxis = pre-configurazione costante dei bit di marcia/sicurezza della command word (template)
   // - Ackerror = reset degli errori del driver dovuti a problemi elettromeccanici irrisolti del motore (non efficace quando tali problemi restano rilevati dal driver) 
   // - HWIDSTW = identificatore hw riferimento telegramma per invio setpoint (parola di comando STW1)
   //   - tipo: HW_IO/HW_ANY
   //   - Sfruttare suggerimenti campo (CTRL + Spazio) per settare in modo simbolico!
   // - HWIDZSW = identificatore hw riferimento telegramma per ricezione actual value (parola di stato ZSW1)
   // 
   // Attenzione: per simulare funzionamento è necessario istanziare un simulatore di interfaccia PROFINet in grado di ricevere e trasmettere word (meglio usare gli Oggetti Tecnologici (come proposto nella network successiva) a fini successivi)
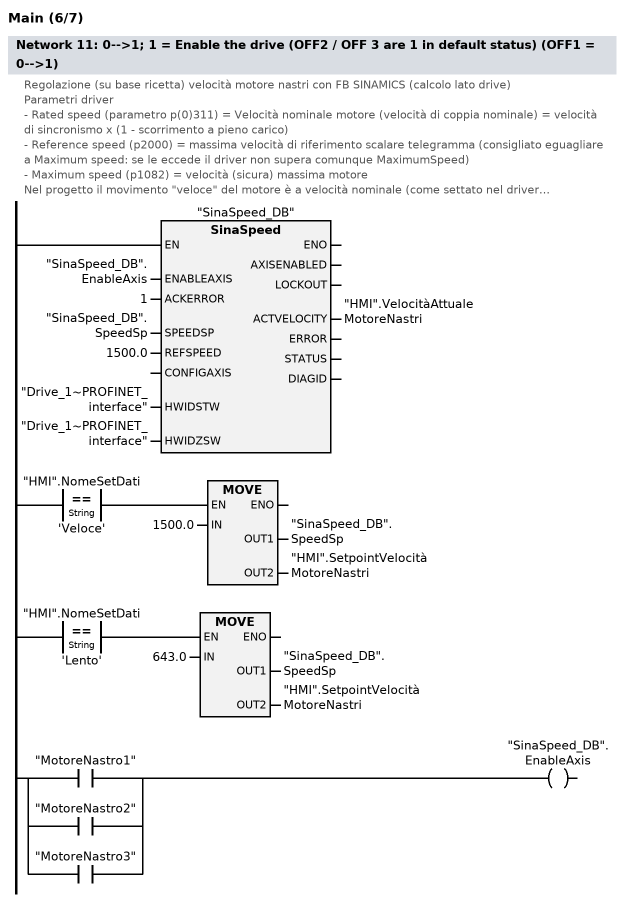
   "SinaSpeed_DB"(EnableAxis := "SinaSpeed_DB".EnableAxis,   // SinaSpeed
                  AckError := 1,
                  SpeedSp := "SinaSpeed_DB".SpeedSp,
                  RefSpeed := 1500.0,
                  HWIDSTW := "Drive_1~PROFINET_interface",
                  HWIDZSW := "Drive_1~PROFINET_interface",
                  ActVelocity => "HMI".VelocitàAttualeMotoreNastri);
   IF "HMI".NomeSetDati = 'Veloce' THEN
       "SinaSpeed_DB".SpeedSp := 1500.0;
       "HMI".SetpointVelocitàMotoreNastri := 1500.0;
   END_IF;
   IF "HMI".NomeSetDati = 'Lento' THEN
       "SinaSpeed_DB".SpeedSp := 643.0;
       "HMI".SetpointVelocitàMotoreNastri := 643.0;
   END_IF;
   "SinaSpeed_DB".EnableAxis := "MotoreNastro1" OR "MotoreNastro2" OR "MotoreNastro3";
END_REGION

REGION Network 12
   // Regolazione (su base ricetta) velocità motore nastri con Technology MC_MoveVelocity (calcolo lato PLC, comunicazione astratta con standard PLCOpen per garantire compatibilità con più costruttori di driver)
   // 
   // Configurazione Oggetto Tecnologico TO_SpeedAxis (in assenza, TO_PositioningAxis):
   // - DRIVE: PROFIdrive
   // - SIMULATION: Simulate drive and encoder
   // - PROFIdrive DATA CONNECTION: Drive
   // - PROFIdrive Drive: Drive.Telegram…
   //   - (sempre necessario telegramma che supporti lettura encoder con TO_PositioningAxis, a meno che l’encoder non sia collegato direttamente al plc)
   //   - (non necessario indicare a fini simulativi)
   // - ENCODER CONNECTION: PROFINET/PROFIBUS
   // - ENCODER DATA CONNECTION: encoder
   //   - (non necessario indicare a fini simulativi)
   // - Dynamics > General Maximum velocity as driver
   // 
   // 
   // Parametri speciali:
   // - Current (velocity) to ignore setpoint and keep actual velocity
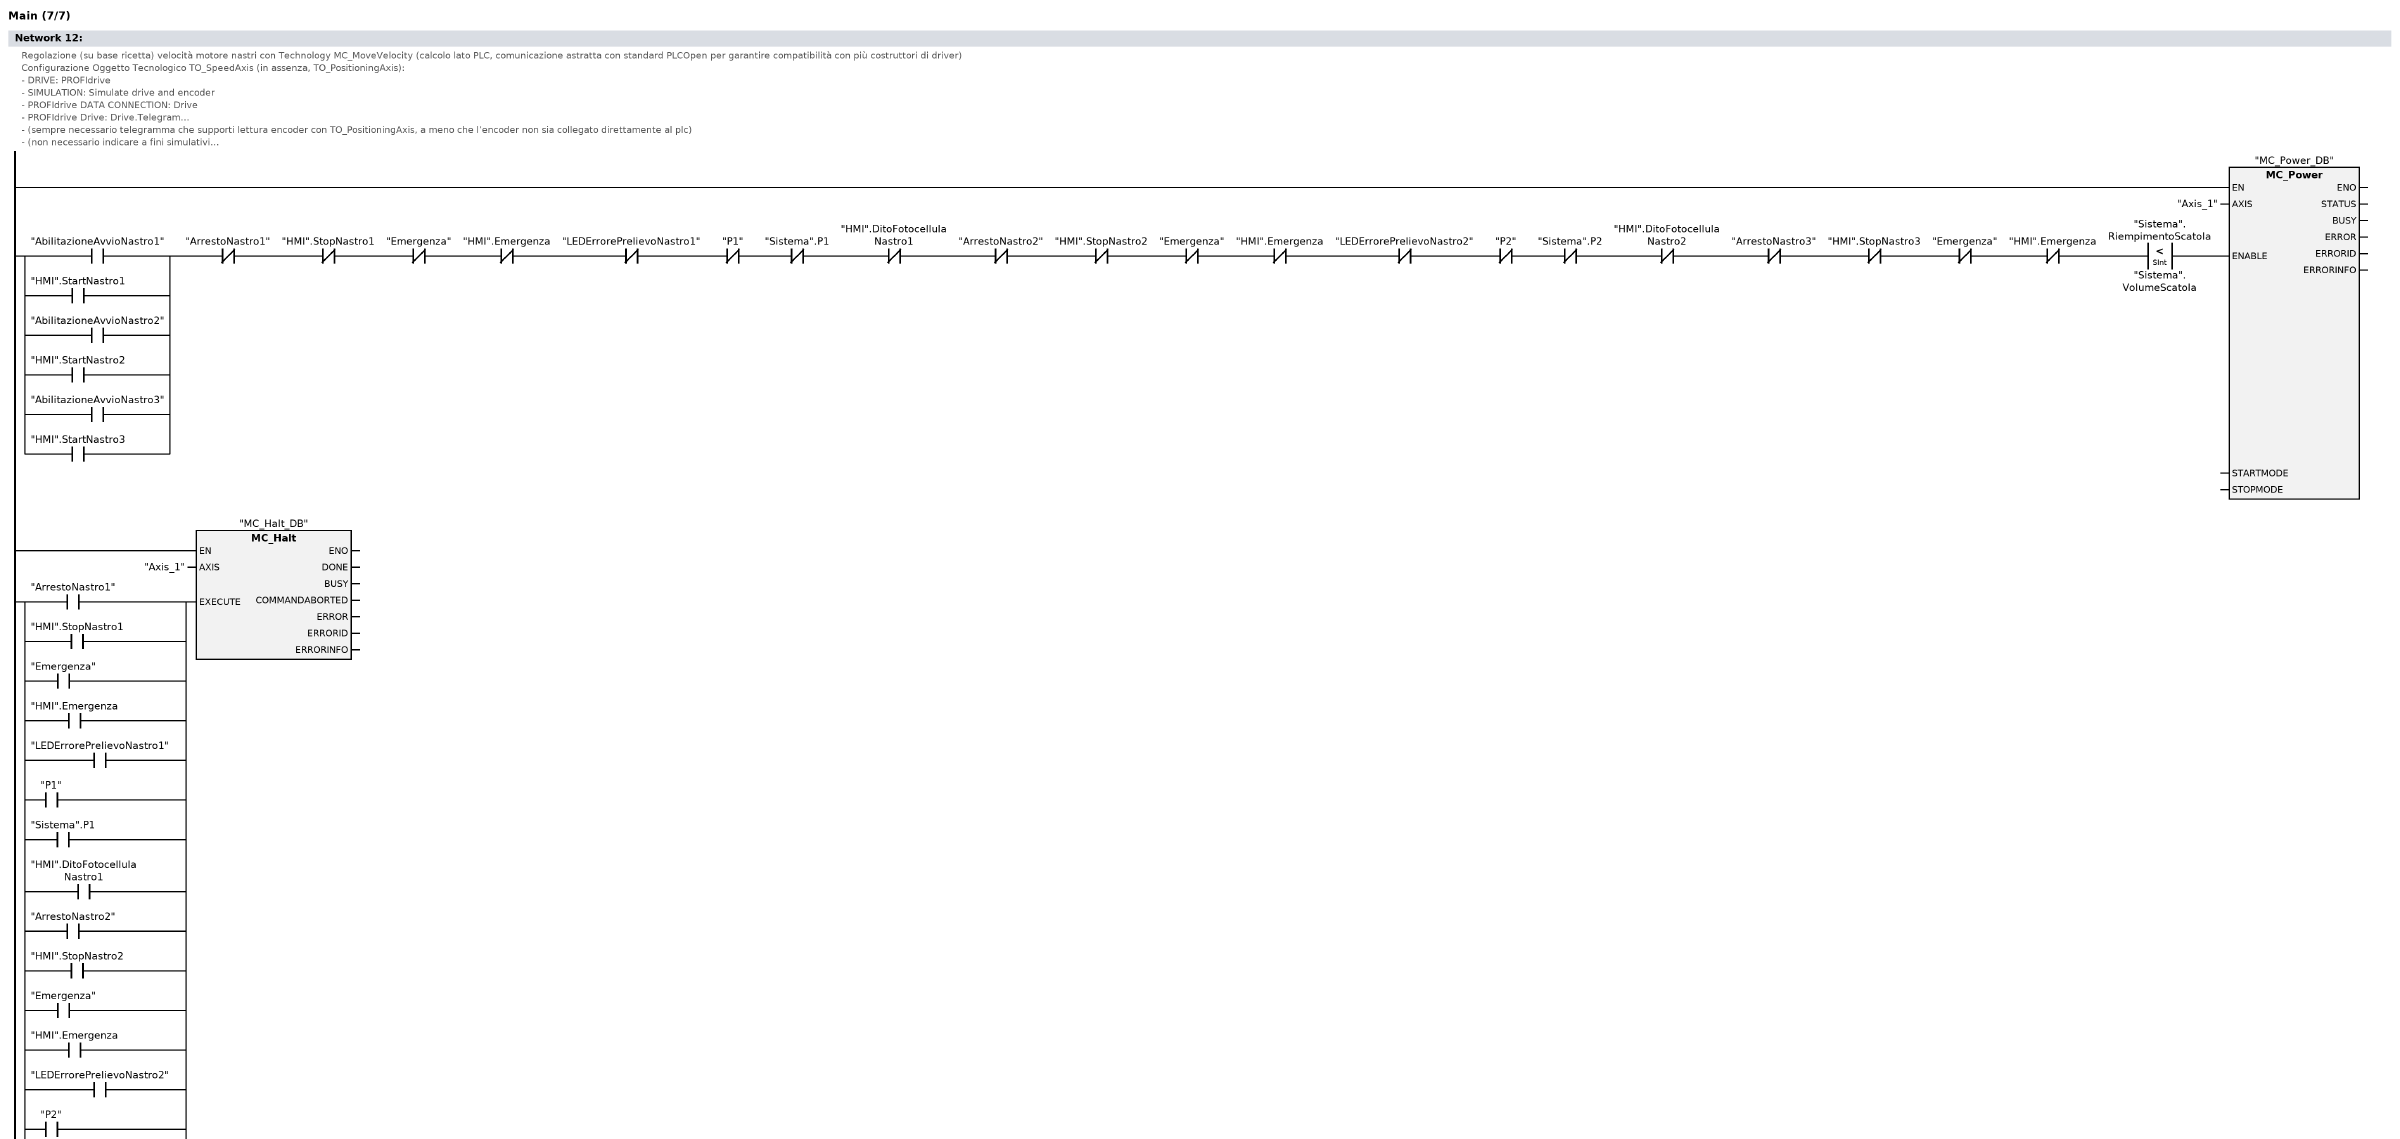
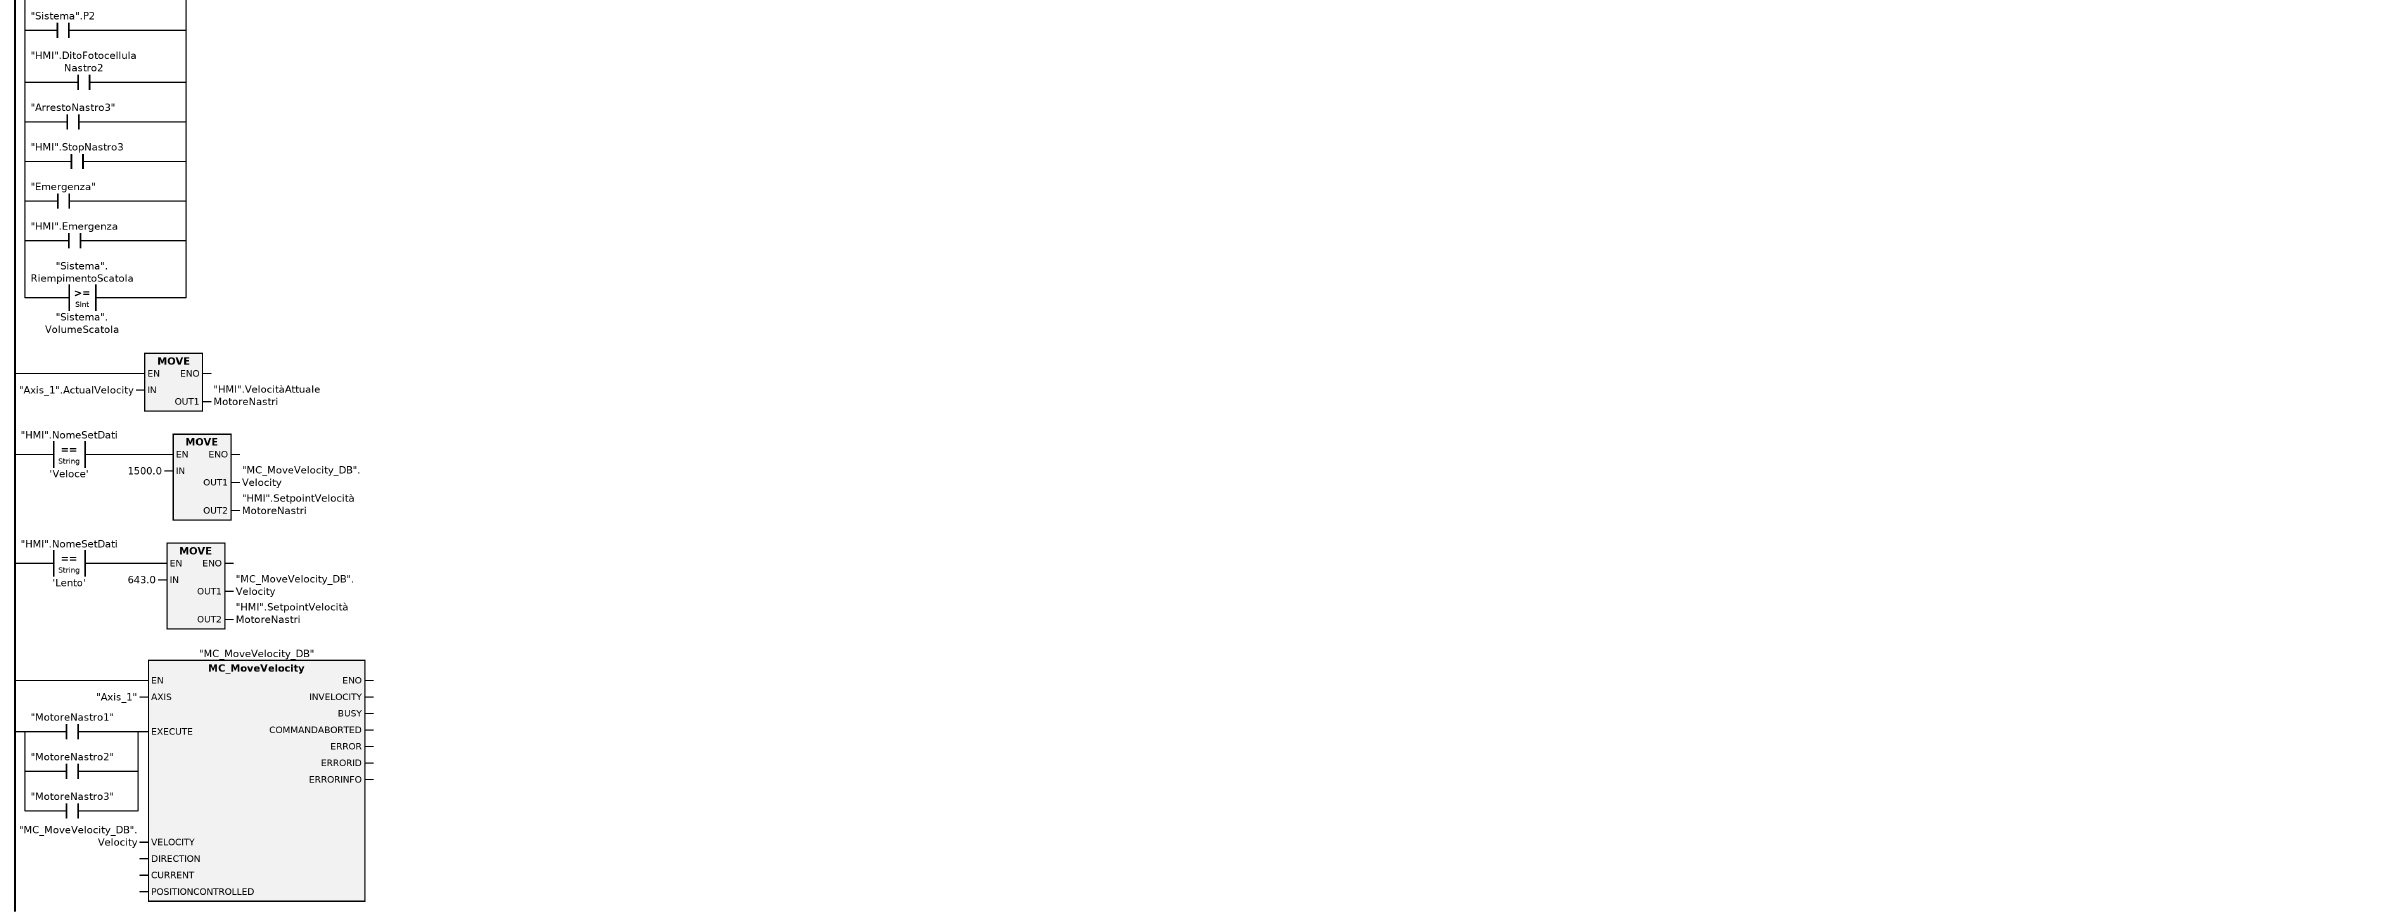
   "MC_Power_DB"(Axis := "Axis_1",   // MC_Power
                 Enable := ("AbilitazioneAvvioNastro1" OR "HMI".StartNastro1 OR "AbilitazioneAvvioNastro2" OR "HMI".StartNastro2 OR "AbilitazioneAvvioNastro3" OR "HMI".StartNastro3) AND NOT "ArrestoNastro1" AND NOT "HMI".StopNastro1 AND NOT "Emergenza" AND NOT "HMI".Emergenza AND NOT "LEDErrorePrelievoNastro1" AND NOT "P1" AND NOT "Sistema".P1 AND NOT "HMI".DitoFotocellulaNastro1 AND NOT "ArrestoNastro2" AND NOT "HMI".StopNastro2 AND NOT "Emergenza" AND NOT "HMI".Emergenza AND NOT "LEDErrorePrelievoNastro2" AND NOT "P2" AND NOT "Sistema".P2 AND NOT "HMI".DitoFotocellulaNastro2 AND NOT "ArrestoNastro3" AND NOT "HMI".StopNastro3 AND NOT "Emergenza" AND NOT "HMI".Emergenza AND ("Sistema".RiempimentoScatola < "Sistema".VolumeScatola));
   "MC_Halt_DB"(Axis := "Axis_1",   // MC_Halt
                Execute := "ArrestoNastro1" OR "HMI".StopNastro1 OR "Emergenza" OR "HMI".Emergenza OR "LEDErrorePrelievoNastro1" OR "P1" OR "Sistema".P1 OR "HMI".DitoFotocellulaNastro1 OR "ArrestoNastro2" OR "HMI".StopNastro2 OR "Emergenza" OR "HMI".Emergenza OR "LEDErrorePrelievoNastro2" OR "P2" OR "Sistema".P2 OR "HMI".DitoFotocellulaNastro2 OR "ArrestoNastro3" OR "HMI".StopNastro3 OR "Emergenza" OR "HMI".Emergenza OR ("Sistema".RiempimentoScatola >= "Sistema".VolumeScatola));
   "HMI".VelocitàAttualeMotoreNastri := "Axis_1".ActualVelocity;
   IF "HMI".NomeSetDati = 'Veloce' THEN
       "MC_MoveVelocity_DB".Velocity := 1500.0;
       "HMI".SetpointVelocitàMotoreNastri := 1500.0;
   END_IF;
   IF "HMI".NomeSetDati = 'Lento' THEN
       "MC_MoveVelocity_DB".Velocity := 643.0;
       "HMI".SetpointVelocitàMotoreNastri := 643.0;
   END_IF;
   "MC_MoveVelocity_DB"(Axis := "Axis_1",   // MC_MoveVelocity
                        Execute := "MotoreNastro1" OR "MotoreNastro2" OR "MotoreNastro3",
                        Velocity := "MC_MoveVelocity_DB".Velocity);
END_REGION
END_ORGANIZATION_BLOCK

(* ===== HMI "HMI_RT_1" =====
system functions are stored by id; their names below are inferred from use
connection "HMI_Collegamento_1": ETHERNET, SMART_S7_1200_OMS

HMI tags "Tabella delle variabili standard"
   "Variabile_Numero di pagina" : UInt, internal
   "Sistema_RiempimentoScatola" : SInt = PLC Sistema.RiempimentoScatola, 100 ms
   "Robot_DB_PosizioneAttuale" : SInt = PLC Robot_DB.PosizioneAttuale, 100 ms
   "HMI_StartNastro3" : Bool = PLC HMI.StartNastro3, 100 ms
   "HMI_StopNastro3" : Bool = PLC HMI.StopNastro3, 100 ms
   "HMI_StartNastro1" : Bool = PLC HMI.StartNastro1, 100 ms
   "HMI_StopNastro1" : Bool = PLC HMI.StopNastro1, 100 ms
   "HMI_StartNastro2" : Bool = PLC HMI.StartNastro2, 100 ms
   "HMI_StopNastro2" : Bool = PLC HMI.StopNastro2, 100 ms
   "LEDErrorePrelievoNastro1" : Bool = PLC LEDErrorePrelievoNastro1 AT %Q0.3, 100 ms
   "LEDErrorePrelievoNastro2" : Bool = PLC LEDErrorePrelievoNastro2 AT %Q1.1, 100 ms
   "HMI_Emergenza" : Bool = PLC HMI.Emergenza, 100 ms
   "HMI_DitoFotocellulaNastro1" : Bool = PLC HMI.DitoFotocellulaNastro1, 100 ms
   "HMI_DitoFotocellulaNastro2" : Bool = PLC HMI.DitoFotocellulaNastro2, 100 ms
   "HMI_CaricamentoPezzoNastro1" : Bool = PLC HMI.CaricamentoPezzoNastro1, 100 ms
   "HMI_CaricamentoPezzoNastro2" : Bool = PLC HMI.CaricamentoPezzoNastro2, 100 ms
   "LEDLavorazione" : Bool = PLC LEDLavorazione AT %Q0.1, 100 ms
   "LEDRiposo" : Bool = PLC LEDRiposo AT %Q0.2, 100 ms
   "HMI_Posizione2PinzaAperta" : Bool = PLC HMI.Posizione2PinzaAperta, 100 ms
   "HMI_Posizione2PinzaChiusa" : Bool = PLC HMI.Posizione2PinzaChiusa, 100 ms
   "HMI_Posizione1PinzaChiusa" : Bool = PLC HMI.Posizione1PinzaChiusa, 100 ms
   "HMI_Posizione1PinzaAperta" : Bool = PLC HMI.Posizione1PinzaAperta, 100 ms
   "HMI_Posizione3PinzaAperta" : Bool = PLC HMI.Posizione3PinzaAperta, 100 ms
   "HMI_Posizione3PinzaChiusa" : Bool = PLC HMI.Posizione3PinzaChiusa, 100 ms
   "Sistema_P1" : Bool = PLC Sistema.P1, 100 ms
   "Sistema_P2" : Bool = PLC Sistema.P2, 100 ms
   "IndiceSegnalazioni" : Int = PLC IndiceSegnalazioni AT %MW100, 100 ms
   "SetDatiSistema_DurataTrasportoNastri" : Time = PLC SetDatiSistema.DurataTrasportoNastri, 100 ms
   "SetDatiSistema_DurataSpostamentoRobot" : Time = PLC SetDatiSistema.DurataSpostamentoRobot, 100 ms
   "SetDatiSistema_VolumeScatola" : SInt = PLC SetDatiSistema.VolumeScatola, 100 ms
   "TPNastro3_ET" : Time = PLC TPNastro3.ET, 100 ms
   "TPNastro1_ET" : Time = PLC TPNastro1.ET, 100 ms
   "TPNastro2_ET" : Time = PLC TPNastro2.ET, 100 ms
   "HMI_IndiceRicetta" : Int = PLC HMI.IndiceRicetta, 100 ms
   "HMI_NomeSetDati" : String[254] = PLC HMI.NomeSetDati, 100 ms
   "TPSostituzioneScatola_Q" : Bool = PLC TPSostituzioneScatola.Q, 100 ms
   "HMI_VisibilitàPezzoNastro3Lento" : Bool = PLC HMI.VisibilitàPezzoNastro3Lento, 100 ms
   "HMI_VisibilitàPezzoNastro3Veloce" : Bool = PLC HMI.VisibilitàPezzoNastro3Veloce, 100 ms
   "HMI_VisibilitàPezzoNastro1Lento" : Bool = PLC HMI.VisibilitàPezzoNastro1Lento, 100 ms
   "HMI_VisibilitàPezzoNastro1Veloce" : Bool = PLC HMI.VisibilitàPezzoNastro1Veloce, 100 ms
   "HMI_VisibilitàPezzoNastro2Lento" : Bool = PLC HMI.VisibilitàPezzoNastro2Lento, 100 ms
   "HMI_VisibilitàPezzoNastro2Veloce" : Bool = PLC HMI.VisibilitàPezzoNastro2Veloce, 100 ms
   "HMI_SetpointVelocitàMotoreNastri" : Real = PLC HMI.SetpointVelocitàMotoreNastri, 1 s
   "HMI_VelocitàAttualeMotoreNastri" : Real = PLC HMI.VelocitàAttualeMotoreNastri, 1 s

discrete alarms
   1: 'Errore Prelievo Nastro 1 - Tentativi in corso...', class Warnings, trigger "IndiceSegnalazioni" bit 0
   2: 'Errore Prelievo Nastro 2 - Tentativi in corso...', class Warnings, trigger "IndiceSegnalazioni" bit 1

text list "Elenco testi_Nome della pagina": 1 'Pagina base'; 2 'Gestione utenti'

recipe "Sistema": DurataTrasportoNastri <- "SetDatiSistema_DurataTrasportoNastri", DurataSpostamentoRobot <- "SetDatiSistema_DurataSpostamentoRobot", VolumeScatola <- "SetDatiSistema_VolumeScatola"

Template "Modello_1" 800x480
   Button "Esci" at 1,42 size 55x39; TextOff 'Esci'; PictureOff "ExitRuntime_KTP900_Basic_PN_TR"; PictureOn "ExitRuntime_KTP900_Basic_PN_TR"
      on Release: StopRuntime(0)
   SymbolicIOField "Pagina_campo_IO_simbolico" at 69,7 size 624x26; TextOff '0'; TextOn '1'; TextList "Elenco testi_Nome della pagina"
      ProcessValue <- "Variabile_Numero di pagina"
      on Change: ActivateScreenByNumber("Variabile_Numero di pagina", 0)
   DateTimeField "HmiScreenItemData" at 695,20 size 105x20
   DateTimeField "HmiScreenItemData_1" at 695,0 size 105x20
   GraphicView "Logo" at 0,0 size 67x40; Picture "Logo di HMI_1"

screen "Processo" 800x480, template "Modello_1"
   on GenerateScreen: SetTag("Variabile_Numero di pagina", 1)
   GraphicView "Vista grafica_6" at 469,326 size 96x72; Picture "pinza45bottom_1"
      Visibility <- "HMI_Posizione2PinzaAperta"
   Rectangle "Rectangle_1" at 402,149 size 60x60
      Appearance <- "TPSostituzioneScatola_Q"
   GraphicView "Vista grafica_4" at 465,230 size 96x48; Picture "pinza45top"
      Visibility <- "HMI_Posizione1PinzaAperta"
   Circle "Cerchio_2" at 476,131 size 54x54
      Appearance <- "LEDRiposo"
   Circle "Cerchio_1" at 475,72 size 54x54
      Appearance <- "LEDLavorazione"
   GraphicIOField "PlotLight_Round_R_1" at 327,130 size 55x55; PictureOff "PilotLight_Round_R_Off_256c"; PictureOn "PilotLight_Round_R_On_256c"
      ProcessValue <- "LEDErrorePrelievoNastro2"
   GraphicIOField "PlotLight_Round_R" at 327,73 size 55x55; PictureOff "PilotLight_Round_R_Off_256c"; PictureOn "PilotLight_Round_R_On_256c"
      ProcessValue <- "LEDErrorePrelievoNastro1"
   GraphicView "Vista grafica_8" at 18,165 size 132x252; Picture "Grafica_8"
   Button "HmiScreenItemData_1" at 62,42 size 145x39; TextOff 'Gestione utenti'; PictureOff "Navigates to Gestione utenti for KTP900 Basic+ PN 17.0.0.0"; PictureOn "Navigates to Gestione utenti for KTP900 Basic+ PN 17.0.0.0"; Authorization "Gestione utenti"
      on Release: ActivateScreen("Gestione utenti", 0)
   GraphicView "Vista grafica_1" at 137,239 size 135x85; Picture "InvertedRetractedPusher"
   GraphicView "Vista grafica_2" at 567,151 size 144x93; Picture "InvertedRetractedPusher"
   GraphicView "Vista grafica_3" at 567,360 size 143x91; Picture "RetractedPusher"
   Button "FB_SlowForward_Round" at 666,151 size 50x50; TextOff 'Text'; PictureOff "FB_SlowForward_Round_Released_256c"; PictureOn "FB_SlowForward_Round_Pressed_256c"
      on Click: SetBit("HMI_StartNastro1"); ResetBit("HMI_StopNastro1")
   Button "FB_SlowForward_Round_1" at 665,406 size 50x50; TextOff 'Text'; PictureOff "FB_SlowForward_Round_Released_256c"; PictureOn "FB_SlowForward_Round_Pressed_256c"
      on Click: SetBit("HMI_StartNastro2"); ResetBit("HMI_StopNastro2")
   Button "FB_SlowForward_Round_2" at 227,239 size 50x50; TextOff 'Text'; PictureOff "FB_SlowForward_Round_Released_256c"; PictureOn "FB_SlowForward_Round_Pressed_256c"
      on Click: SetBit("HMI_StartNastro3"); ResetBit("HMI_StopNastro3")
   Button "FB_Stop_Round" at 563,406 size 50x50; TextOff 'Text'; PictureOff "FB_Stop_Round_Released_256c"; PictureOn "FB_Stop_Round_Pressed_256c"
      on Press: SetBit("HMI_StopNastro2"); ResetBit("HMI_StartNastro2")
   Button "FB_Stop_Round_1" at 562,151 size 50x50; TextOff 'Text'; PictureOff "FB_Stop_Round_Released_256c"; PictureOn "FB_Stop_Round_Pressed_256c"
      on Press: SetBit("HMI_StopNastro1"); ResetBit("HMI_StartNastro1")
   Button "FB_Stop_Round_2" at 132,239 size 50x50; TextOff 'Text'; PictureOff "FB_Stop_Round_Released_256c"; PictureOn "FB_Stop_Round_Pressed_256c"
      on Press: SetBit("HMI_StopNastro3"); ResetBit("HMI_StartNastro3")
   GraphicView "Vista grafica_9" at 393,354 size 71x104; Picture "PinzaBottom"
      Visibility <- "Robot_DB_PosizioneAttuale"
   GraphicView "Vista grafica_10" at 657,203 size 76x40; Picture "Cjstiel"
      HorizontalMovement <- "TPNastro1_ET"
      Visibility <- "HMI_VisibilitàPezzoNastro1Veloce"
   GraphicView "Vista grafica_11" at 661,360 size 76x40; Picture "Cjstiel"
      HorizontalMovement <- "TPNastro2_ET"
      Visibility <- "HMI_VisibilitàPezzoNastro2Veloce"
   GraphicView "Vista grafica_12" at 212,285 size 76x40; Picture "Cjstiel"
      HorizontalMovement <- "TPNastro3_ET"
      Visibility <- "HMI_VisibilitàPezzoNastro3Veloce"
   TextField "Casella di testo_1" at 475,51 size 56x20; Text 'Sistema'
   TextField "Casella di testo_2" at 334,51 size 41x20; Text 'Errori'
   Button "FB_Plus_Round" at 693,246 size 50x50; TextOff 'Text'; PictureOff "FB_Plus_Round_Released_256c"; PictureOn "FB_Plus_Round_Pressed_256c"
      on Press: SetBit("HMI_CaricamentoPezzoNastro1")
      on Release: ResetBit("HMI_CaricamentoPezzoNastro1")
   Button "FB_Cross_Round" at 570,246 size 50x50; TextOff 'Text'; PictureOff "FB_Cross_Round_Released_256c"; PictureOn "FB_Cross_Round_Pressed_256c"
      on Press: SetBit("HMI_DitoFotocellulaNastro1")
      on Release: ResetBit("HMI_DitoFotocellulaNastro1")
   Button "FB_Plus_Round_1" at 694,308 size 50x50; TextOff 'Text'; PictureOff "FB_Plus_Round_Released_256c"; PictureOn "FB_Plus_Round_Pressed_256c"
      on Release: ResetBit("HMI_CaricamentoPezzoNastro2")
      on Press: SetBit("HMI_CaricamentoPezzoNastro2")
   Button "FB_Cross_Round_1" at 570,309 size 50x50; TextOff 'Text'; PictureOff "FB_Cross_Round_Released_256c"; PictureOn "FB_Cross_Round_Pressed_256c"
      on Release: ResetBit("HMI_DitoFotocellulaNastro2")
      on Press: SetBit("HMI_DitoFotocellulaNastro2")
   TextField "Casella di testo_3" at 329,86 size 48x36; Text 'Nastro 1'
   TextField "Casella di testo_4" at 330,143 size 52x36; Text 'Nastro 2'
   TextField "Casella di testo_6" at 480,137 size 45x36; Text 'A riposo'
   TextField "Casella di testo_5" at 478,77 size 48x36; Text 'In marcia'
   TextField "Casella di testo_7" at 406,151 size 52x52; Text 'Sostitu zione scatola'
   TextField "Casella di testo_8" at 394,51 size 76x20; Text 'Emergenza'
   TextField "Casella di testo_9" at 568,131 size 35x20; Text 'Stop'
   TextField "Casella di testo_10" at 570,456 size 35x20; Text 'Stop'
   TextField "Casella di testo_11" at 140,216 size 35x20; Text 'Stop'
   TextField "Casella di testo_12" at 229,216 size 39x20; Text 'Start'
   TextField "Casella di testo_13" at 671,456 size 39x20; Text 'Start'
   TextField "Casella di testo_14" at 670,131 size 39x20; Text 'Start'
   TextField "Casella di testo_15" at 722,154 size 62x42; Text 'NASTRO 1'
   TextField "Casella di testo_16" at 726,411 size 62x42; Text 'NASTRO 2'
   TextField "Casella di testo_17" at 176,330 size 74x26; Text 'NASTRO 3'
   TextField "Casella di testo_18" at 746,245 size 46x52; Text 'Carica mento pezzo'
   TextField "Casella di testo_19" at 749,307 size 46x52; Text 'Carica mento pezzo'
   TextField "Casella di testo_20" at 622,245 size 72x52; Text 'Dito sulla fotocellula'
   TextField "Casella di testo_21" at 622,307 size 72x52; Text 'Dito sulla fotocellula'
   GraphicView "Vista grafica_16" at 56,314 size 61x39; Picture "Cjstiel"
      Visibility <- "Sistema_RiempimentoScatola"
   GraphicView "Vista grafica_17" at 55,272 size 61x39; Picture "Cjstiel"
      Visibility <- "Sistema_RiempimentoScatola"
   GraphicView "Vista grafica_18" at 55,229 size 61x42; Picture "Cjstiel"
      Visibility <- "Sistema_RiempimentoScatola"
   Button "Pulsante_1" at 548,41 size 107x39; TextOff 'Segnalazioni'; Authorization "Accesso segnalazioni"
      on Click: ActivateScreen("Segnalazioni", 0)
   Button "Pulsante_2" at 667,41 size 128x39; TextOff 'Gestione ricette'; Authorization "Gestione ricette"
      on Click: ActivateScreen("Gestione ricette", 0)
   Switch "Pushbutton_Emergency" at 397,74 size 68x66; CaptionText 'Switch'; TextOff '0'; TextOn '1'; PictureOn "Pushbutton_Emergency_On_256c"; PictureOff "Pushbutton_Emergency_Off_256c"
      ProcessValue <- "HMI_Emergenza"
      on SwitchOn: SetBit("HMI_Emergenza")
      on SwitchOff: ResetBit("HMI_Emergenza")
   GraphicView "Vista grafica_19" at 548,203 size 76x40; Picture "Cjstiel"
      Visibility <- "Sistema_P1"
   GraphicView "Vista grafica_20" at 559,360 size 76x40; Picture "Cjstiel"
      Visibility <- "Sistema_P2"
   GraphicView "Vista grafica_15" at 464,230 size 96x48; Picture "pinzaChiusaBottom2"
      Visibility <- "HMI_Posizione1PinzaChiusa"
   GraphicView "Vista grafica_13" at 462,314 size 98x82; Picture "pinzaChiusaBottom"
      Visibility <- "HMI_Posizione2PinzaChiusa"
   GraphicView "Vista grafica_5" at 278,282 size 96x48; Picture "pinza"
      Visibility <- "HMI_Posizione3PinzaAperta"
   GraphicView "Vista grafica_14" at 280,261 size 96x82; Picture "pinzaChiusa"
      Visibility <- "HMI_Posizione3PinzaChiusa"
   GraphicView "Vista grafica_7" at 361,236 size 132x133; Picture "Grafica_4"
   GraphicView "Vista grafica_21" at 53,297 size 61x39; Picture "Cjstiel"
      Visibility <- "Sistema_RiempimentoScatola"
   GraphicView "Vista grafica_22" at 53,250 size 61x39; Picture "Cjstiel"
      Visibility <- "Sistema_RiempimentoScatola"
   GraphicView "Vista grafica_23" at 50,272 size 61x39; Picture "Cjstiel"
      Visibility <- "Sistema_RiempimentoScatola"
   GraphicView "Vista grafica_24" at 212,286 size 76x40; Picture "Cjstiel"
      HorizontalMovement <- "TPNastro3_ET"
      Visibility <- "HMI_VisibilitàPezzoNastro3Lento"
   GraphicView "Vista grafica_25" at 657,203 size 76x40; Picture "Cjstiel"
      HorizontalMovement <- "TPNastro1_ET"
      Visibility <- "HMI_VisibilitàPezzoNastro1Lento"
   GraphicView "Vista grafica_26" at 662,360 size 76x40; Picture "Cjstiel"
      HorizontalMovement <- "TPNastro2_ET"
      Visibility <- "HMI_VisibilitàPezzoNastro2Lento"
   IOField "I/O field_1" at 172,110 size 96x32; FormatPattern s9999.999
      ProcessValue <- "HMI_SetpointVelocitàMotoreNastri"
   IOField "I/O field_2" at 171,167 size 96x32; FormatPattern s9999.999
      ProcessValue <- "HMI_VelocitàAttualeMotoreNastri"
   TextField "Text field_1" at 141,88 size 157x20; Text 'Setpoint velocità nastri'
   TextField "Text field_2" at 141,144 size 150x20; Text 'Velocità attuale nastri'

screen "Gestione utenti" 800x480, template "Modello_1"
   on GenerateScreen: SetTag("Variabile_Numero di pagina", 2)
   UserView "HmiScreenItemData" at 0,89 size 799x390
   Button "Indietro" at 57,41 size 159x47; TextOff 'Indietro'
      on Release: ActivateScreen("Processo", 0)
   Button "Pulsante_1" at 273,44 size 192x32; TextOff 'Segnalazioni'; Authorization "Accesso segnalazioni"
      on Click: ActivateScreen("Segnalazioni", 0)
   Button "Pulsante_2" at 510,44 size 192x32; TextOff 'Gestione ricette'; Authorization "Gestione ricette"
      on Click: ActivateScreen("Gestione ricette", 0)

screen "Segnalazioni" 800x480
   AlarmView "Vista segnalazioni_1" at 0,0 size 799x326; ColumnTextClassName 'Classe'
   Button "Pulsante_1" at 4,434 size 192x32; TextOff 'Gestione utenti'; Authorization "Gestione utenti"
      on Click: ActivateScreen("Gestione utenti", 0)
   Button "Pulsante_2" at 206,434 size 192x32; TextOff 'Processo'
      on Click: ActivateScreen("Processo", 0)
   Button "Pulsante_3" at 407,434 size 192x32; TextOff 'Gestione ricette'; Authorization "Gestione ricette"
      on Click: ActivateScreen("Gestione ricette", 0)
   Button "Pulsante_4" at 650,434 size 147x32; TextOff 'Reset segnalazioni'
      on Click: function_e14cd482(0)

screen "Gestione ricette" 800x480
   RecipeView "Vista ricette_1" at 0,0 size 799x407; Recipe "Sistema"; Tag4RecipeNumber "HMI_IndiceRicetta"; Tag4DataRecord "HMI_NomeSetDati"
   Button "Pulsante_1" at 26,423 size 192x32; TextOff 'Gestione utenti'; Authorization "Gestione utenti"
      on Click: ActivateScreen("Gestione utenti", 0)
   Button "Pulsante_2" at 269,423 size 192x32; TextOff 'Processo'
      on Click: ActivateScreen("Processo", 0)
   Button "Pulsante_3" at 506,423 size 192x32; TextOff 'Segnalazioni'; Authorization "Accesso segnalazioni"
      on Click: ActivateScreen("Segnalazioni", 0)
*)